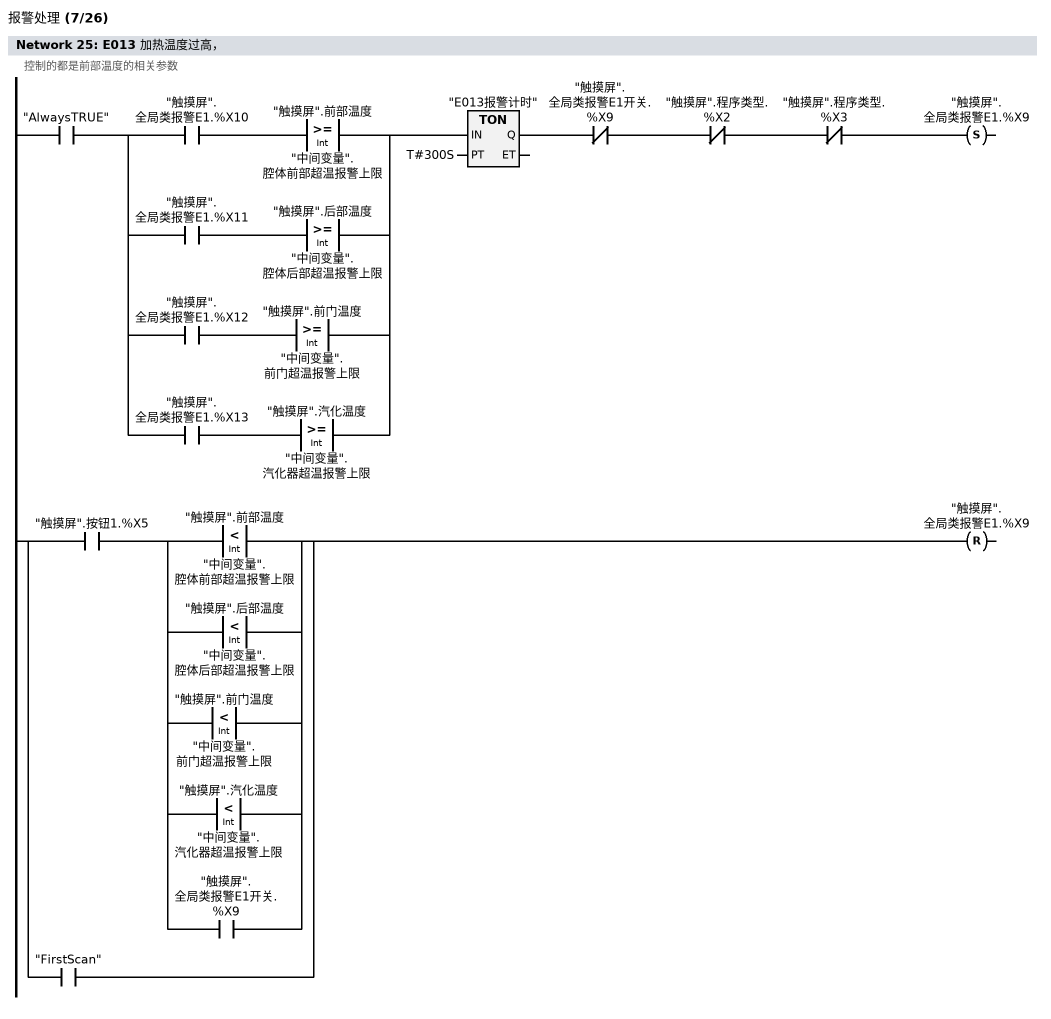
   "E013报警计时".TON(IN := "AlwaysTRUE" AND (("触摸屏".全局类报警E1.%X10 AND ("触摸屏".前部温度 >= "中间变量".腔体前部超温报警上限)) OR ("触摸屏".全局类报警E1.%X11 AND ("触摸屏".后部温度 >= "中间变量".腔体后部超温报警上限)) OR ("触摸屏".全局类报警E1.%X12 AND ("触摸屏".前门温度 >= "中间变量".前门超温报警上限)) OR ("触摸屏".全局类报警E1.%X13 AND ("触摸屏".汽化温度 >= "中间变量".汽化器超温报警上限))),
                  PT := T#300S);
   IF "E013报警计时".Q AND NOT "触摸屏".全局类报警E1开关.%X9 AND NOT "触摸屏".程序类型.%X2 AND NOT "触摸屏".程序类型.%X3 THEN
       "触摸屏".全局类报警E1.%X9 := TRUE;
   END_IF;
   IF ("触摸屏".按钮1.%X5 AND (("触摸屏".前部温度 < "中间变量".腔体前部超温报警上限) OR ("触摸屏".后部温度 < "中间变量".腔体后部超温报警上限) OR ("触摸屏".前门温度 < "中间变量".前门超温报警上限) OR ("触摸屏".汽化温度 < "中间变量".汽化器超温报警上限) OR "触摸屏".全局类报警E1开关.%X9)) OR "FirstScan" THEN
       "触摸屏".全局类报警E1.%X9 := FALSE;
   END_IF;
END_REGION

REGION Network 26: E014 加热系统异常，加热系统断电-脱扣器
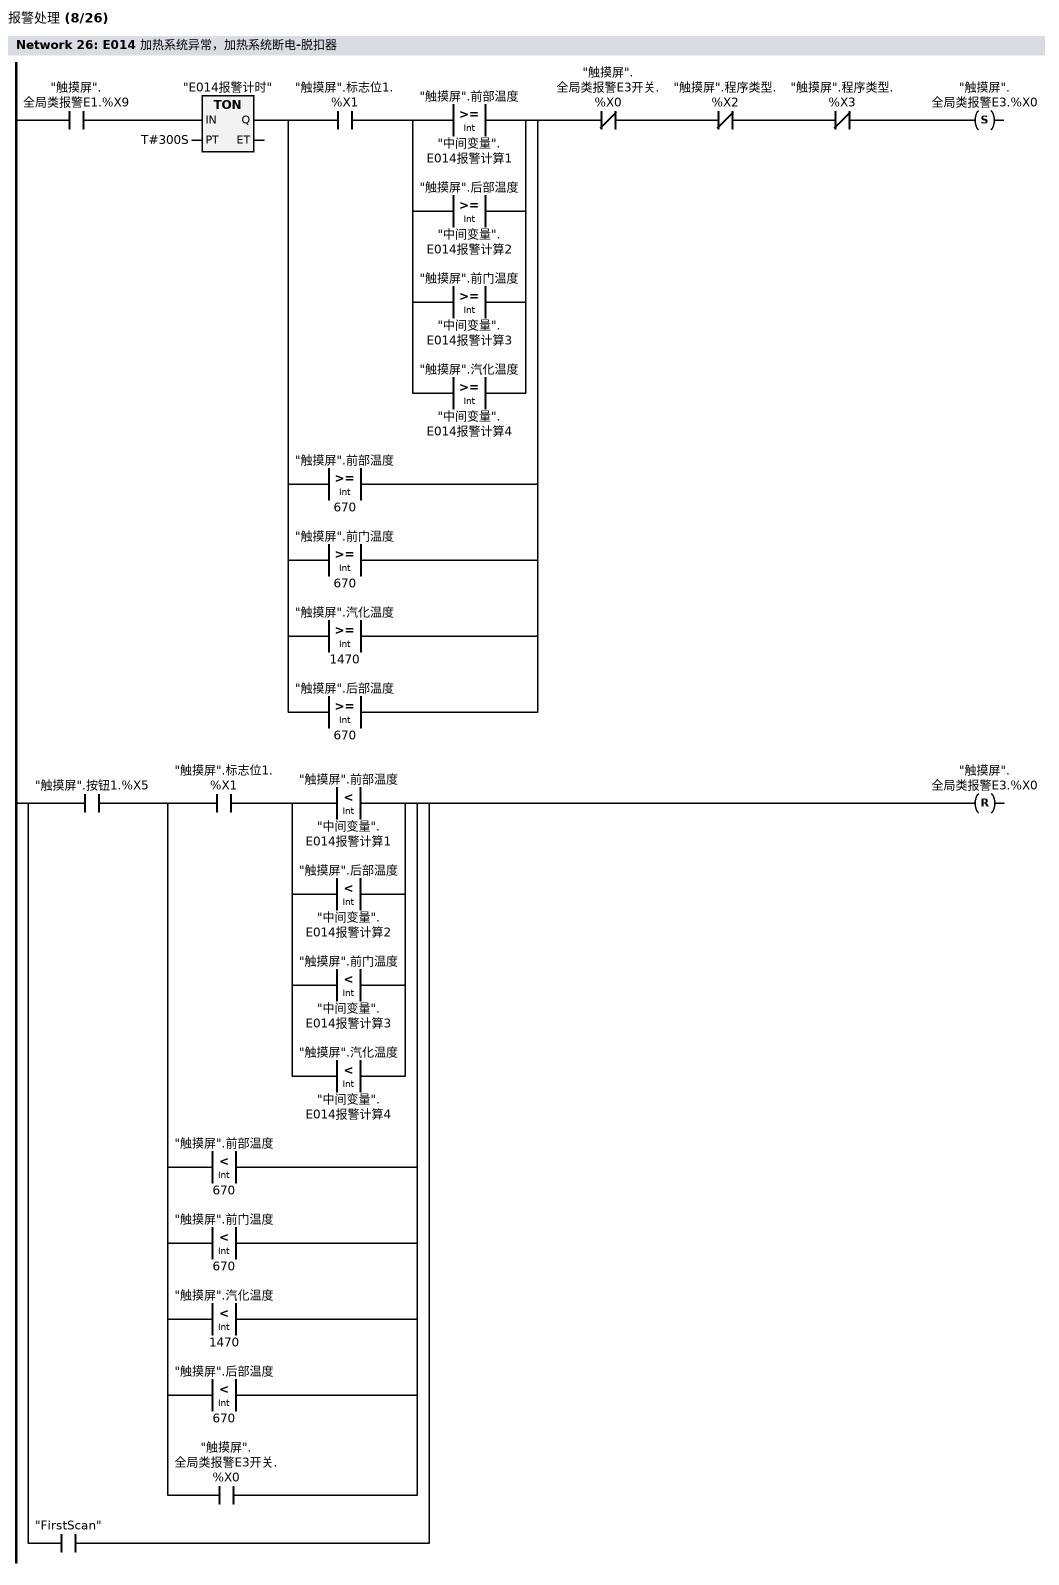
   "E014报警计时".TON(IN := "触摸屏".全局类报警E1.%X9, PT := T#300S);
   IF "E014报警计时".Q AND (("触摸屏".标志位1.%X1 AND (("触摸屏".前部温度 >= "中间变量".E014报警计算1) OR ("触摸屏".后部温度 >= "中间变量".E014报警计算2) OR ("触摸屏".前门温度 >= "中间变量".E014报警计算3) OR ("触摸屏".汽化温度 >= "中间变量".E014报警计算4))) OR ("触摸屏".前部温度 >= 670) OR ("触摸屏".前门温度 >= 670) OR ("触摸屏".汽化温度 >= 1470) OR ("触摸屏".后部温度 >= 670)) AND NOT "触摸屏".全局类报警E3开关.%X0 AND NOT "触摸屏".程序类型.%X2 AND NOT "触摸屏".程序类型.%X3 THEN
       "触摸屏".全局类报警E3.%X0 := TRUE;
   END_IF;
   IF ("触摸屏".按钮1.%X5 AND (("触摸屏".标志位1.%X1 AND (("触摸屏".前部温度 < "中间变量".E014报警计算1) OR ("触摸屏".后部温度 < "中间变量".E014报警计算2) OR ("触摸屏".前门温度 < "中间变量".E014报警计算3) OR ("触摸屏".汽化温度 < "中间变量".E014报警计算4))) OR ("触摸屏".前部温度 < 670) OR ("触摸屏".前门温度 < 670) OR ("触摸屏".汽化温度 < 1470) OR ("触摸屏".后部温度 < 670) OR "触摸屏".全局类报警E3开关.%X0)) OR "FirstScan" THEN
       "触摸屏".全局类报警E3.%X0 := FALSE;
   END_IF;
END_REGION

REGION Network 27: E015 腔体前部超温
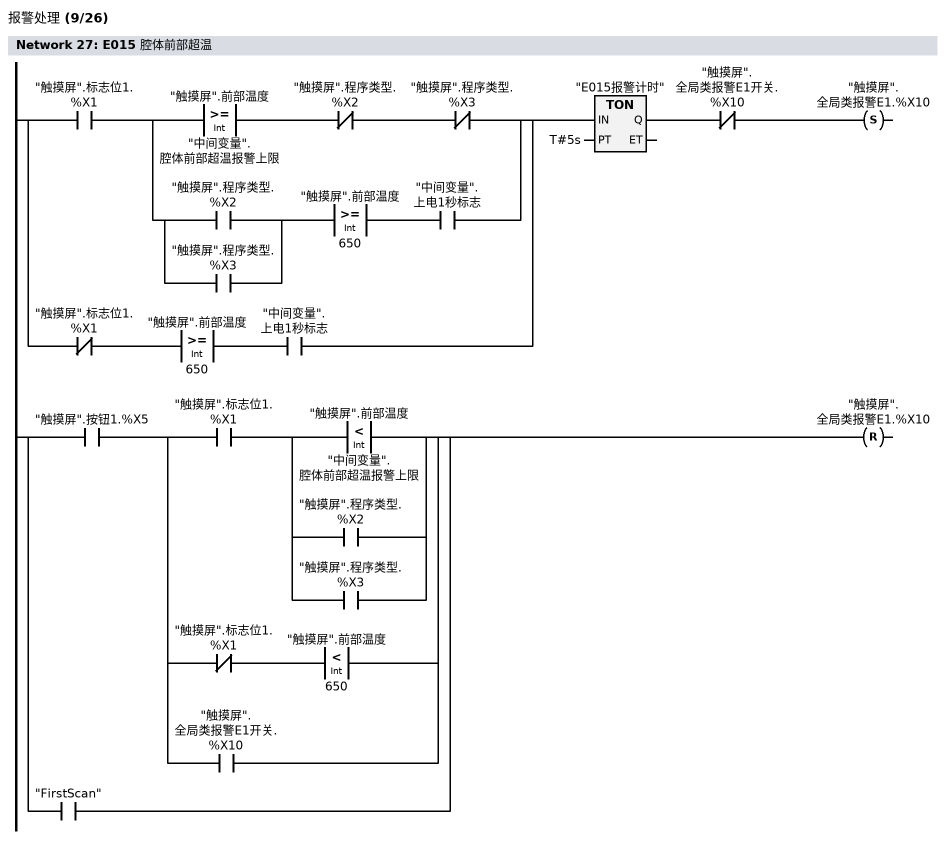
   "E015报警计时".TON(IN := ("触摸屏".标志位1.%X1 AND ((("触摸屏".前部温度 >= "中间变量".腔体前部超温报警上限) AND NOT "触摸屏".程序类型.%X2 AND NOT "触摸屏".程序类型.%X3) OR (("触摸屏".程序类型.%X2 OR "触摸屏".程序类型.%X3) AND ("触摸屏".前部温度 >= 650) AND "中间变量".上电1秒标志))) OR (NOT "触摸屏".标志位1.%X1 AND ("触摸屏".前部温度 >= 650) AND "中间变量".上电1秒标志),
                  PT := T#5s);
   IF "E015报警计时".Q AND NOT "触摸屏".全局类报警E1开关.%X10 THEN "触摸屏".全局类报警E1.%X10 := TRUE; END_IF;
   IF ("触摸屏".按钮1.%X5 AND (("触摸屏".标志位1.%X1 AND (("触摸屏".前部温度 < "中间变量".腔体前部超温报警上限) OR "触摸屏".程序类型.%X2 OR "触摸屏".程序类型.%X3)) OR (NOT "触摸屏".标志位1.%X1 AND ("触摸屏".前部温度 < 650)) OR "触摸屏".全局类报警E1开关.%X10)) OR "FirstScan" THEN
       "触摸屏".全局类报警E1.%X10 := FALSE;
   END_IF;
END_REGION

REGION Network 28: E016 腔体后部超温
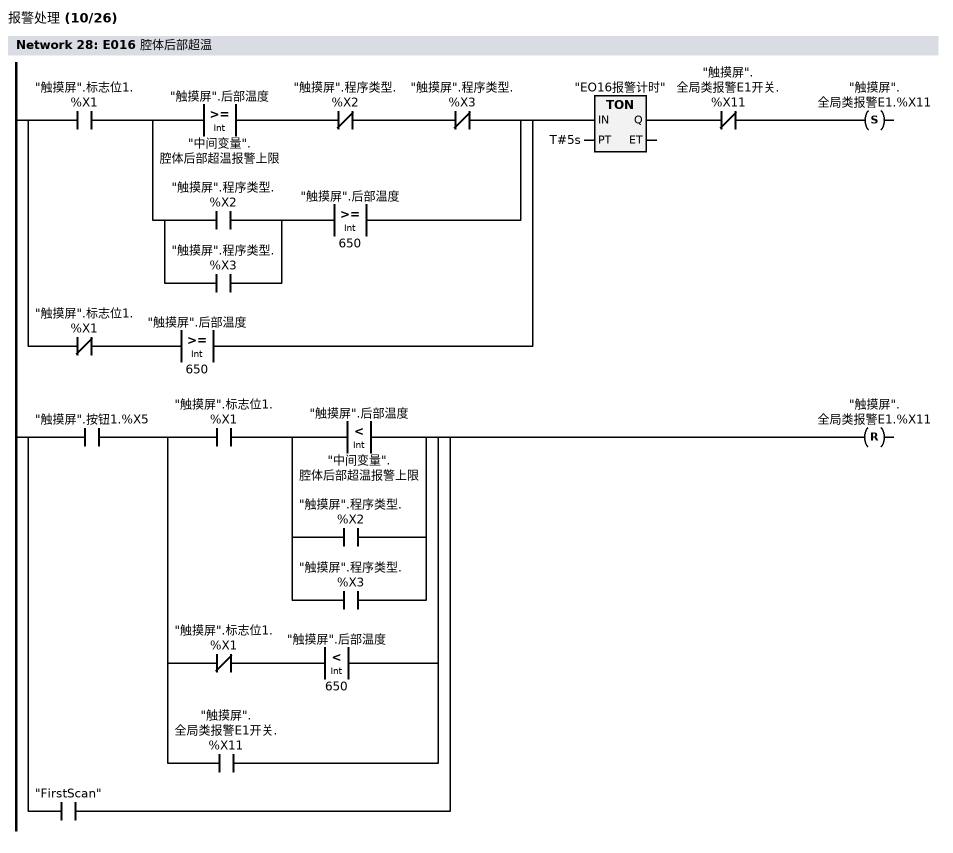
   "EO16报警计时".TON(IN := ("触摸屏".标志位1.%X1 AND ((("触摸屏".后部温度 >= "中间变量".腔体后部超温报警上限) AND NOT "触摸屏".程序类型.%X2 AND NOT "触摸屏".程序类型.%X3) OR (("触摸屏".程序类型.%X2 OR "触摸屏".程序类型.%X3) AND ("触摸屏".后部温度 >= 650)))) OR (NOT "触摸屏".标志位1.%X1 AND ("触摸屏".后部温度 >= 650)),
                  PT := T#5s);
   IF "EO16报警计时".Q AND NOT "触摸屏".全局类报警E1开关.%X11 THEN "触摸屏".全局类报警E1.%X11 := TRUE; END_IF;
   IF ("触摸屏".按钮1.%X5 AND (("触摸屏".标志位1.%X1 AND (("触摸屏".后部温度 < "中间变量".腔体后部超温报警上限) OR "触摸屏".程序类型.%X2 OR "触摸屏".程序类型.%X3)) OR (NOT "触摸屏".标志位1.%X1 AND ("触摸屏".后部温度 < 650)) OR "触摸屏".全局类报警E1开关.%X11)) OR "FirstScan" THEN
       "触摸屏".全局类报警E1.%X11 := FALSE;
   END_IF;
END_REGION

REGION Network 29: E017 门超温
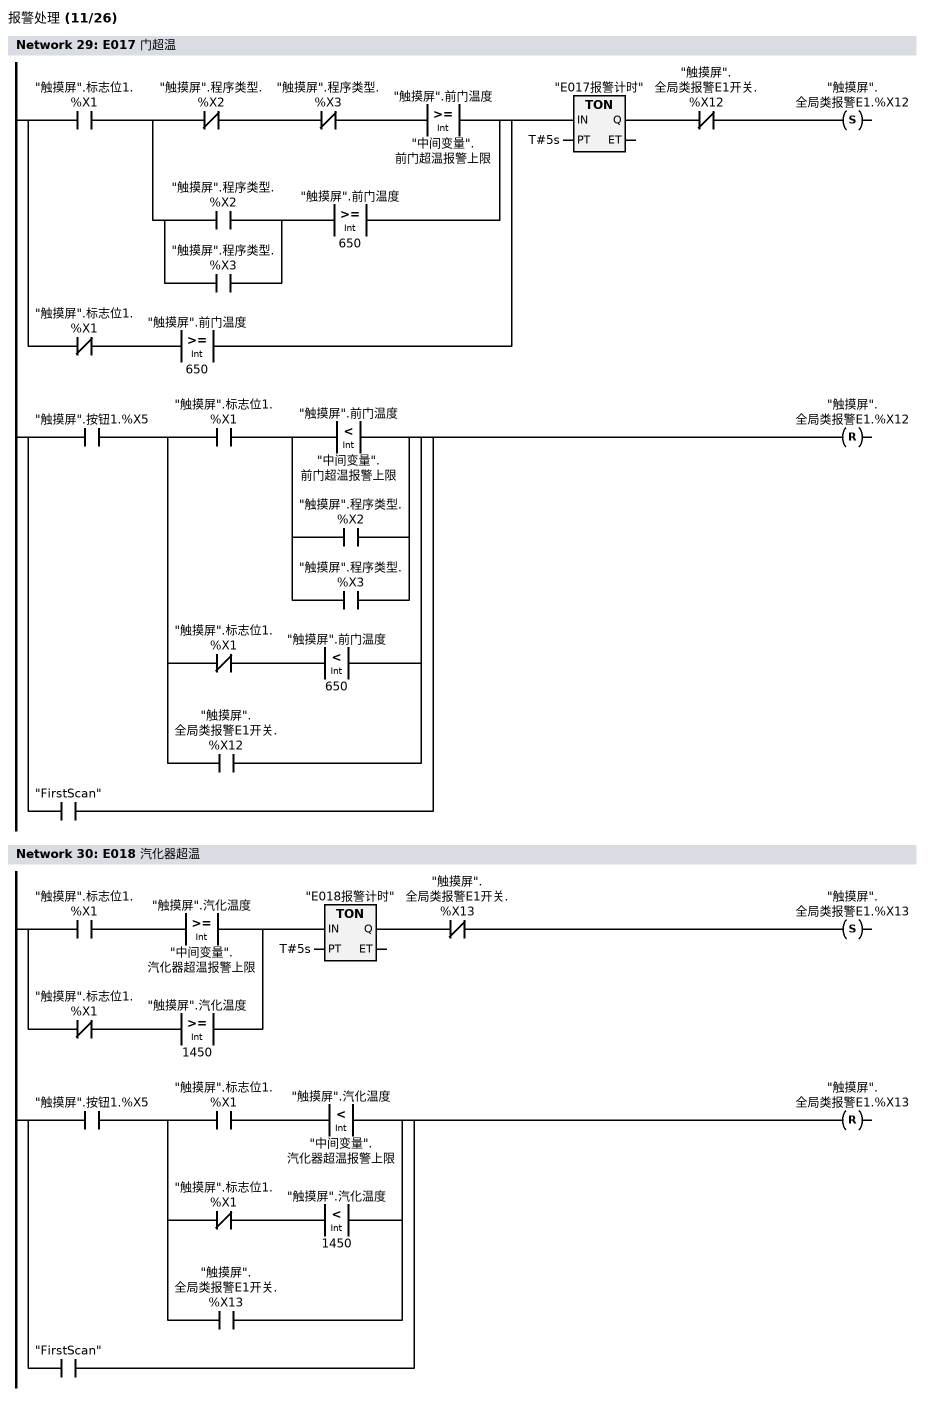
   "E017报警计时".TON(IN := ("触摸屏".标志位1.%X1 AND ((NOT "触摸屏".程序类型.%X2 AND NOT "触摸屏".程序类型.%X3 AND ("触摸屏".前门温度 >= "中间变量".前门超温报警上限)) OR (("触摸屏".程序类型.%X2 OR "触摸屏".程序类型.%X3) AND ("触摸屏".前门温度 >= 650)))) OR (NOT "触摸屏".标志位1.%X1 AND ("触摸屏".前门温度 >= 650)),
                  PT := T#5s);
   IF "E017报警计时".Q AND NOT "触摸屏".全局类报警E1开关.%X12 THEN "触摸屏".全局类报警E1.%X12 := TRUE; END_IF;
   IF ("触摸屏".按钮1.%X5 AND (("触摸屏".标志位1.%X1 AND (("触摸屏".前门温度 < "中间变量".前门超温报警上限) OR "触摸屏".程序类型.%X2 OR "触摸屏".程序类型.%X3)) OR (NOT "触摸屏".标志位1.%X1 AND ("触摸屏".前门温度 < 650)) OR "触摸屏".全局类报警E1开关.%X12)) OR "FirstScan" THEN
       "触摸屏".全局类报警E1.%X12 := FALSE;
   END_IF;
END_REGION

REGION Network 30: E018 汽化器超温
   "E018报警计时".TON(IN := ("触摸屏".标志位1.%X1 AND ("触摸屏".汽化温度 >= "中间变量".汽化器超温报警上限)) OR (NOT "触摸屏".标志位1.%X1 AND ("触摸屏".汽化温度 >= 1450)),
                  PT := T#5s);
   IF "E018报警计时".Q AND NOT "触摸屏".全局类报警E1开关.%X13 THEN "触摸屏".全局类报警E1.%X13 := TRUE; END_IF;
   IF ("触摸屏".按钮1.%X5 AND (("触摸屏".标志位1.%X1 AND ("触摸屏".汽化温度 < "中间变量".汽化器超温报警上限)) OR (NOT "触摸屏".标志位1.%X1 AND ("触摸屏".汽化温度 < 1450)) OR "触摸屏".全局类报警E1开关.%X13)) OR "FirstScan" THEN
       "触摸屏".全局类报警E1.%X13 := FALSE;
   END_IF;
END_REGION

REGION Network 31: E019 内室温度过高
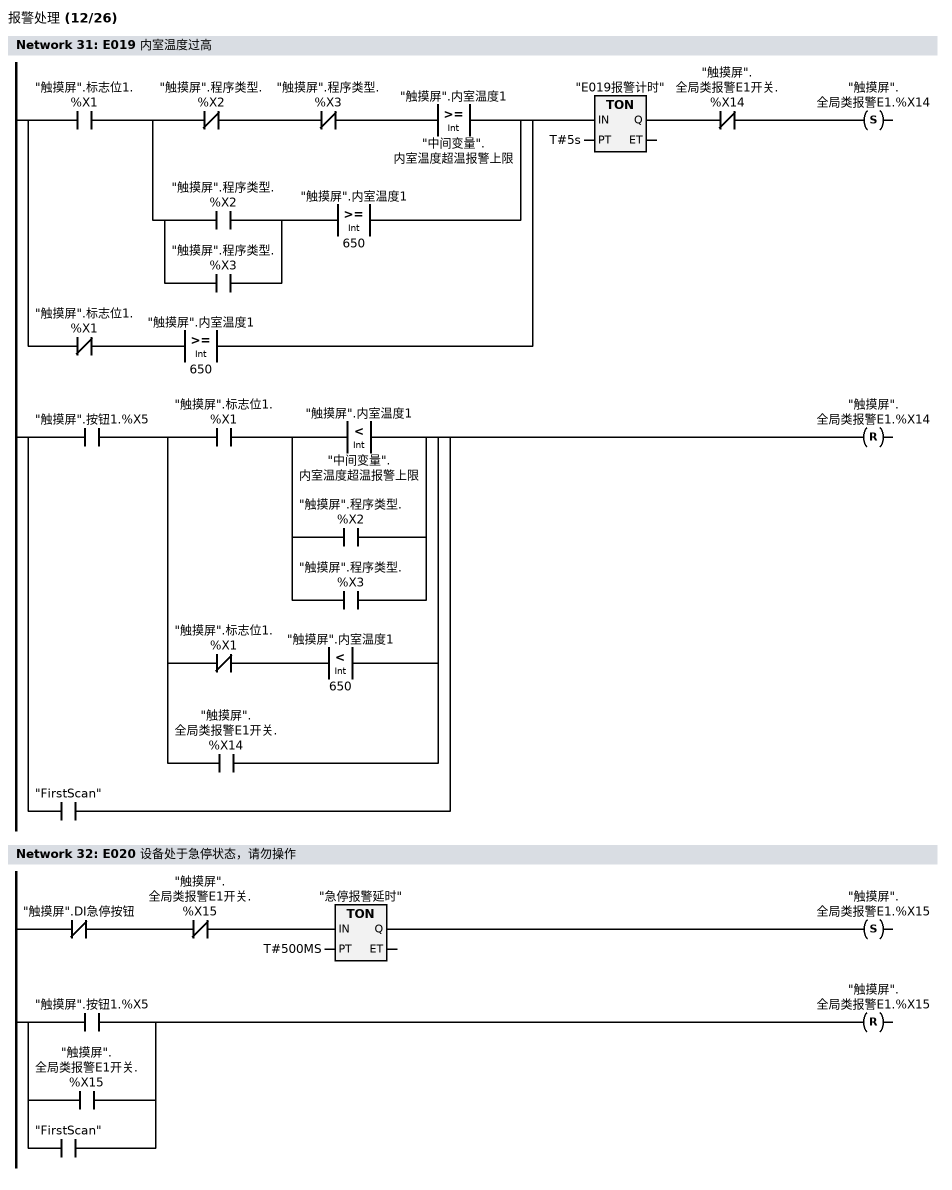
   "E019报警计时".TON(IN := ("触摸屏".标志位1.%X1 AND ((NOT "触摸屏".程序类型.%X2 AND NOT "触摸屏".程序类型.%X3 AND ("触摸屏".内室温度1 >= "中间变量".内室温度超温报警上限)) OR (("触摸屏".程序类型.%X2 OR "触摸屏".程序类型.%X3) AND ("触摸屏".内室温度1 >= 650)))) OR (NOT "触摸屏".标志位1.%X1 AND ("触摸屏".内室温度1 >= 650)),
                  PT := T#5s);
   IF "E019报警计时".Q AND NOT "触摸屏".全局类报警E1开关.%X14 THEN "触摸屏".全局类报警E1.%X14 := TRUE; END_IF;
   IF ("触摸屏".按钮1.%X5 AND (("触摸屏".标志位1.%X1 AND (("触摸屏".内室温度1 < "中间变量".内室温度超温报警上限) OR "触摸屏".程序类型.%X2 OR "触摸屏".程序类型.%X3)) OR (NOT "触摸屏".标志位1.%X1 AND ("触摸屏".内室温度1 < 650)) OR "触摸屏".全局类报警E1开关.%X14)) OR "FirstScan" THEN
       "触摸屏".全局类报警E1.%X14 := FALSE;
   END_IF;
END_REGION

REGION Network 32: E020 设备处于急停状态，请勿操作
   "急停报警延时".TON(IN := NOT "触摸屏".DI急停按钮 AND NOT "触摸屏".全局类报警E1开关.%X15, PT := T#500MS);
   IF "急停报警延时".Q THEN "触摸屏".全局类报警E1.%X15 := TRUE; END_IF;
   IF "触摸屏".按钮1.%X5 OR "触摸屏".全局类报警E1开关.%X15 OR "FirstScan" THEN "触摸屏".全局类报警E1.%X15 := FALSE; END_IF;
END_REGION

REGION Network 33: E021灭菌器与尾气处理器通讯故障
   // 带尾气处理器的设备   通讯超时60秒 我们认为通讯故障
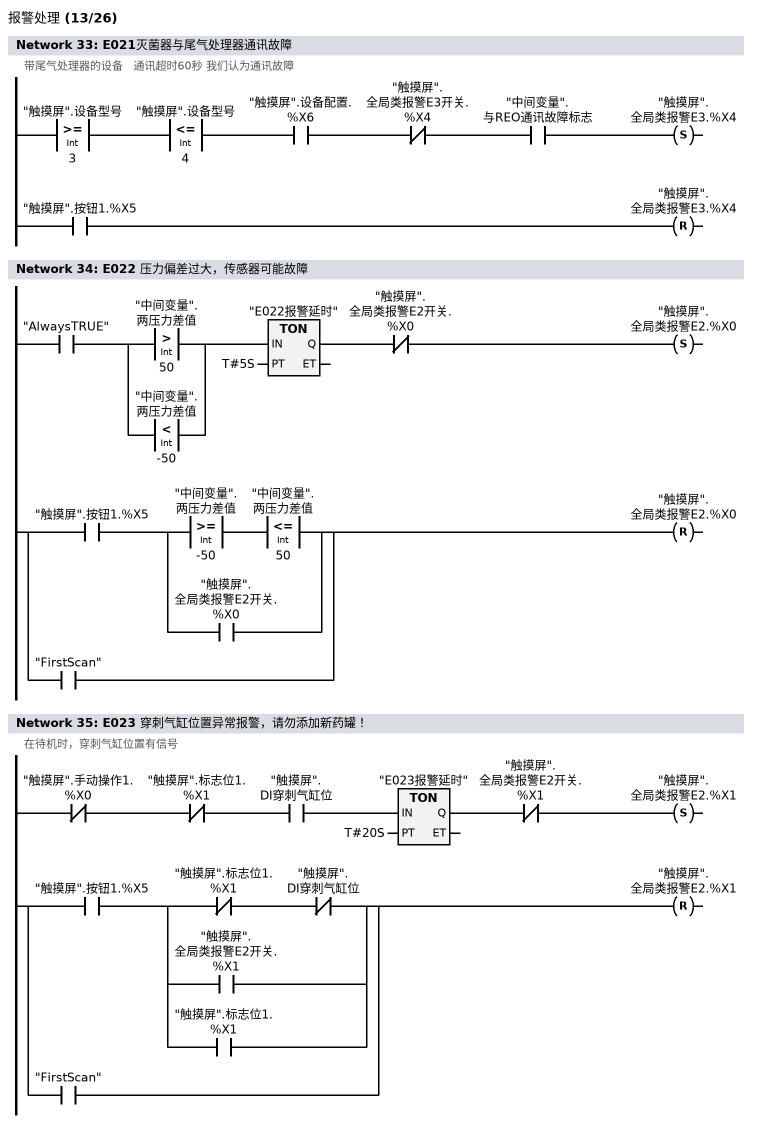
   RUNG wire#powerrail
      { S7_Templates := "SrcType := Int" } GE_Contact(in1 := "触摸屏".设备型号, in2 := 3)
      { S7_Templates := "SrcType := Int" } LE_Contact(in1 := "触摸屏".设备型号, in2 := 4)
      Contact( "触摸屏".设备配置.%X6 )
      I_Contact( "触摸屏".全局类报警E3开关.%X4 )
      Contact( "中间变量".与REO通讯故障标志 )
      S_Coil( "触摸屏".全局类报警E3.%X4 )
   END_RUNG
   RUNG wire#powerrail
      Contact( "触摸屏".按钮1.%X5 )
      R_Coil( "触摸屏".全局类报警E3.%X4 )
   END_RUNG
   // the same network as SCL:
   IF ("触摸屏".设备型号 >= 3) AND ("触摸屏".设备型号 <= 4) AND "触摸屏".设备配置.%X6 AND NOT "触摸屏".全局类报警E3开关.%X4 AND "中间变量".与REO通讯故障标志 THEN
       "触摸屏".全局类报警E3.%X4 := TRUE;
   END_IF;
   IF "触摸屏".按钮1.%X5 THEN "触摸屏".全局类报警E3.%X4 := FALSE; END_IF;
END_REGION

REGION Network 34: E022 压力偏差过大，传感器可能故障
   "E022报警延时".TON(IN := "AlwaysTRUE" AND (("中间变量".两压力差值 > 50) OR ("中间变量".两压力差值 < (-50))), PT := T#5S);
   IF "E022报警延时".Q AND NOT "触摸屏".全局类报警E2开关.%X0 THEN "触摸屏".全局类报警E2.%X0 := TRUE; END_IF;
   IF ("触摸屏".按钮1.%X5 AND ((("中间变量".两压力差值 >= (-50)) AND ("中间变量".两压力差值 <= 50)) OR "触摸屏".全局类报警E2开关.%X0)) OR "FirstScan" THEN
       "触摸屏".全局类报警E2.%X0 := FALSE;
   END_IF;
END_REGION

REGION Network 35: E023 穿刺气缸位置异常报警，请勿添加新药罐！
   // 在待机时，穿刺气缸位置有信号
   "E023报警延时".TON(IN := NOT "触摸屏".手动操作1.%X0 AND NOT "触摸屏".标志位1.%X1 AND "触摸屏".DI穿刺气缸位, PT := T#20S);
   IF "E023报警延时".Q AND NOT "触摸屏".全局类报警E2开关.%X1 THEN "触摸屏".全局类报警E2.%X1 := TRUE; END_IF;
   IF ("触摸屏".按钮1.%X5 AND ((NOT "触摸屏".标志位1.%X1 AND NOT "触摸屏".DI穿刺气缸位) OR "触摸屏".全局类报警E2开关.%X1 OR "触摸屏".标志位1.%X1)) OR "FirstScan" THEN
       "触摸屏".全局类报警E2.%X1 := FALSE;
   END_IF;
END_REGION

REGION Network 36: E024舱体前部温度升温超时
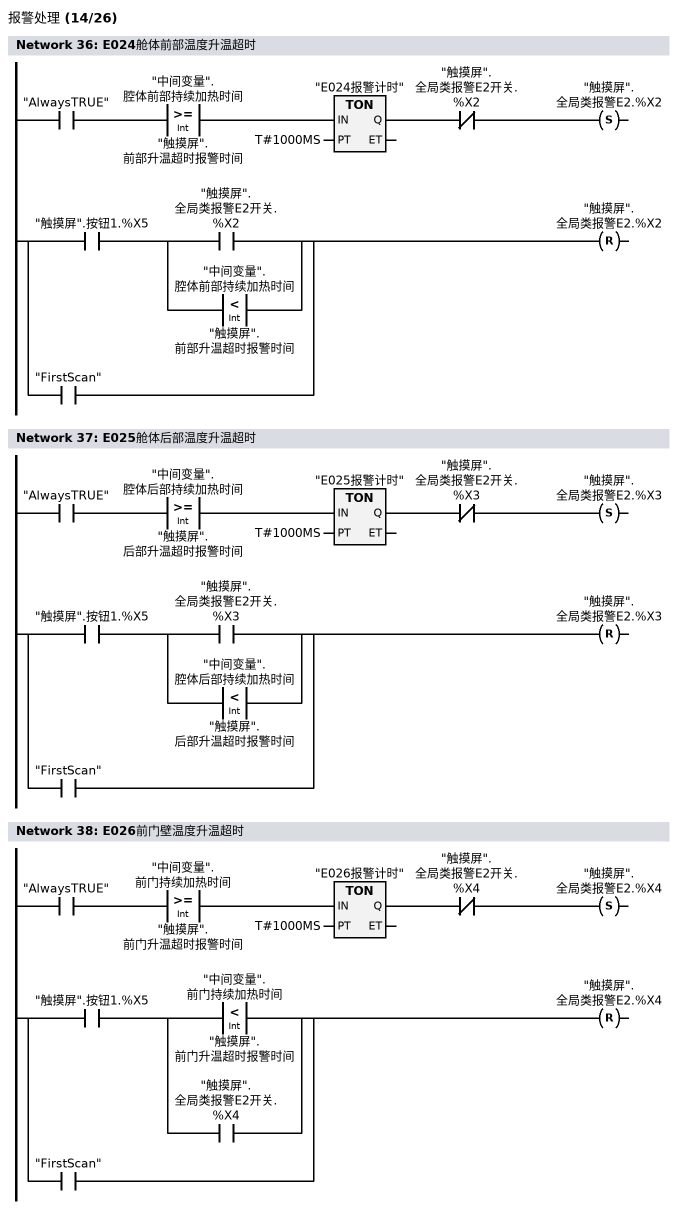
   "E024报警计时".TON(IN := "AlwaysTRUE" AND ("中间变量".腔体前部持续加热时间 >= "触摸屏".前部升温超时报警时间), PT := T#1000MS);
   IF "E024报警计时".Q AND NOT "触摸屏".全局类报警E2开关.%X2 THEN "触摸屏".全局类报警E2.%X2 := TRUE; END_IF;
   IF ("触摸屏".按钮1.%X5 AND ("触摸屏".全局类报警E2开关.%X2 OR ("中间变量".腔体前部持续加热时间 < "触摸屏".前部升温超时报警时间))) OR "FirstScan" THEN
       "触摸屏".全局类报警E2.%X2 := FALSE;
   END_IF;
END_REGION

REGION Network 37: E025舱体后部温度升温超时
   "E025报警计时".TON(IN := "AlwaysTRUE" AND ("中间变量".腔体后部持续加热时间 >= "触摸屏".后部升温超时报警时间), PT := T#1000MS);
   IF "E025报警计时".Q AND NOT "触摸屏".全局类报警E2开关.%X3 THEN "触摸屏".全局类报警E2.%X3 := TRUE; END_IF;
   IF ("触摸屏".按钮1.%X5 AND ("触摸屏".全局类报警E2开关.%X3 OR ("中间变量".腔体后部持续加热时间 < "触摸屏".后部升温超时报警时间))) OR "FirstScan" THEN
       "触摸屏".全局类报警E2.%X3 := FALSE;
   END_IF;
END_REGION

REGION Network 38: E026前门壁温度升温超时
   "E026报警计时".TON(IN := "AlwaysTRUE" AND ("中间变量".前门持续加热时间 >= "触摸屏".前门升温超时报警时间), PT := T#1000MS);
   IF "E026报警计时".Q AND NOT "触摸屏".全局类报警E2开关.%X4 THEN "触摸屏".全局类报警E2.%X4 := TRUE; END_IF;
   IF ("触摸屏".按钮1.%X5 AND (("中间变量".前门持续加热时间 < "触摸屏".前门升温超时报警时间) OR "触摸屏".全局类报警E2开关.%X4)) OR "FirstScan" THEN
       "触摸屏".全局类报警E2.%X4 := FALSE;
   END_IF;
END_REGION

REGION Network 39: E027汽化器温度升温超时
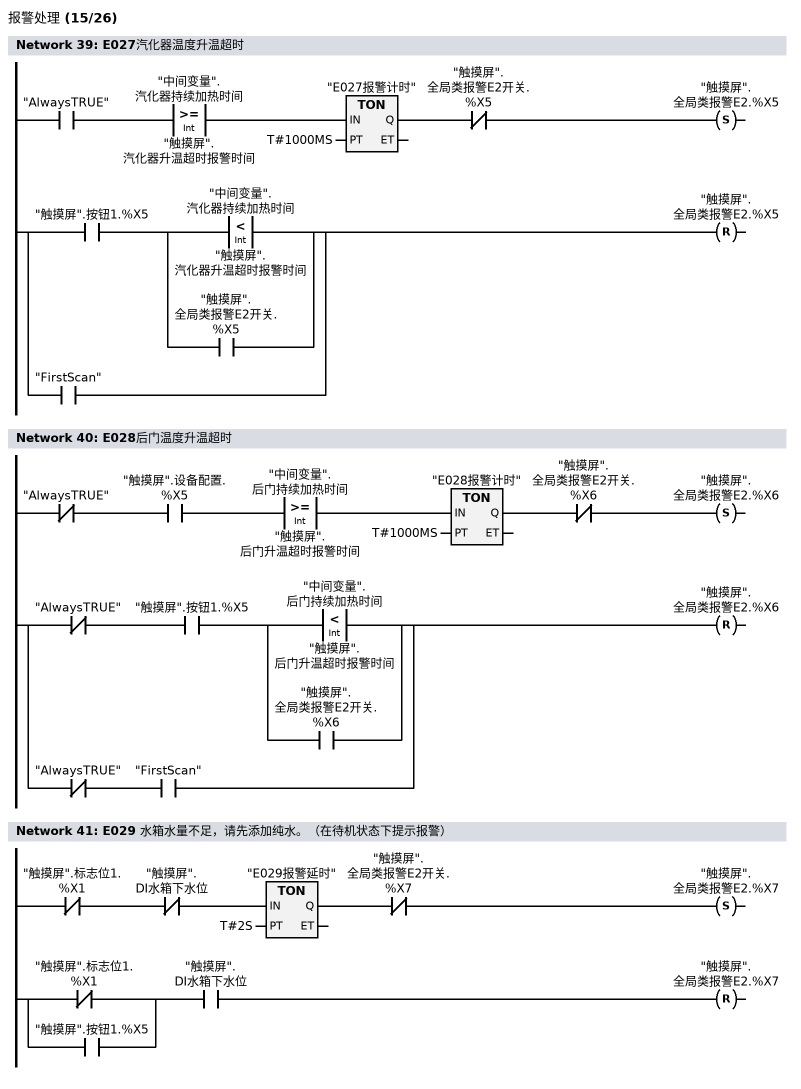
   "E027报警计时".TON(IN := "AlwaysTRUE" AND ("中间变量".汽化器持续加热时间 >= "触摸屏".汽化器升温超时报警时间), PT := T#1000MS);
   IF "E027报警计时".Q AND NOT "触摸屏".全局类报警E2开关.%X5 THEN "触摸屏".全局类报警E2.%X5 := TRUE; END_IF;
   IF ("触摸屏".按钮1.%X5 AND (("中间变量".汽化器持续加热时间 < "触摸屏".汽化器升温超时报警时间) OR "触摸屏".全局类报警E2开关.%X5)) OR "FirstScan" THEN
       "触摸屏".全局类报警E2.%X5 := FALSE;
   END_IF;
END_REGION

REGION Network 40: E028后门温度升温超时
   "E028报警计时".TON(IN := NOT "AlwaysTRUE" AND "触摸屏".设备配置.%X5 AND ("中间变量".后门持续加热时间 >= "触摸屏".后门升温超时报警时间),
                  PT := T#1000MS);
   IF "E028报警计时".Q AND NOT "触摸屏".全局类报警E2开关.%X6 THEN "触摸屏".全局类报警E2.%X6 := TRUE; END_IF;
   IF (NOT "AlwaysTRUE" AND "触摸屏".按钮1.%X5 AND (("中间变量".后门持续加热时间 < "触摸屏".后门升温超时报警时间) OR "触摸屏".全局类报警E2开关.%X6)) OR (NOT "AlwaysTRUE" AND "FirstScan") THEN
       "触摸屏".全局类报警E2.%X6 := FALSE;
   END_IF;
END_REGION

REGION Network 41: E029 水箱水量不足，请先添加纯水。（在待机状态下提示报警）
   "E029报警延时".TON(IN := NOT "触摸屏".标志位1.%X1 AND NOT "触摸屏".DI水箱下水位, PT := T#2S);
   IF "E029报警延时".Q AND NOT "触摸屏".全局类报警E2开关.%X7 THEN "触摸屏".全局类报警E2.%X7 := TRUE; END_IF;
   IF (NOT "触摸屏".标志位1.%X1 OR "触摸屏".按钮1.%X5) AND "触摸屏".DI水箱下水位 THEN "触摸屏".全局类报警E2.%X7 := FALSE; END_IF;
END_REGION

REGION Network 42: E030催化前温度传感器故障！
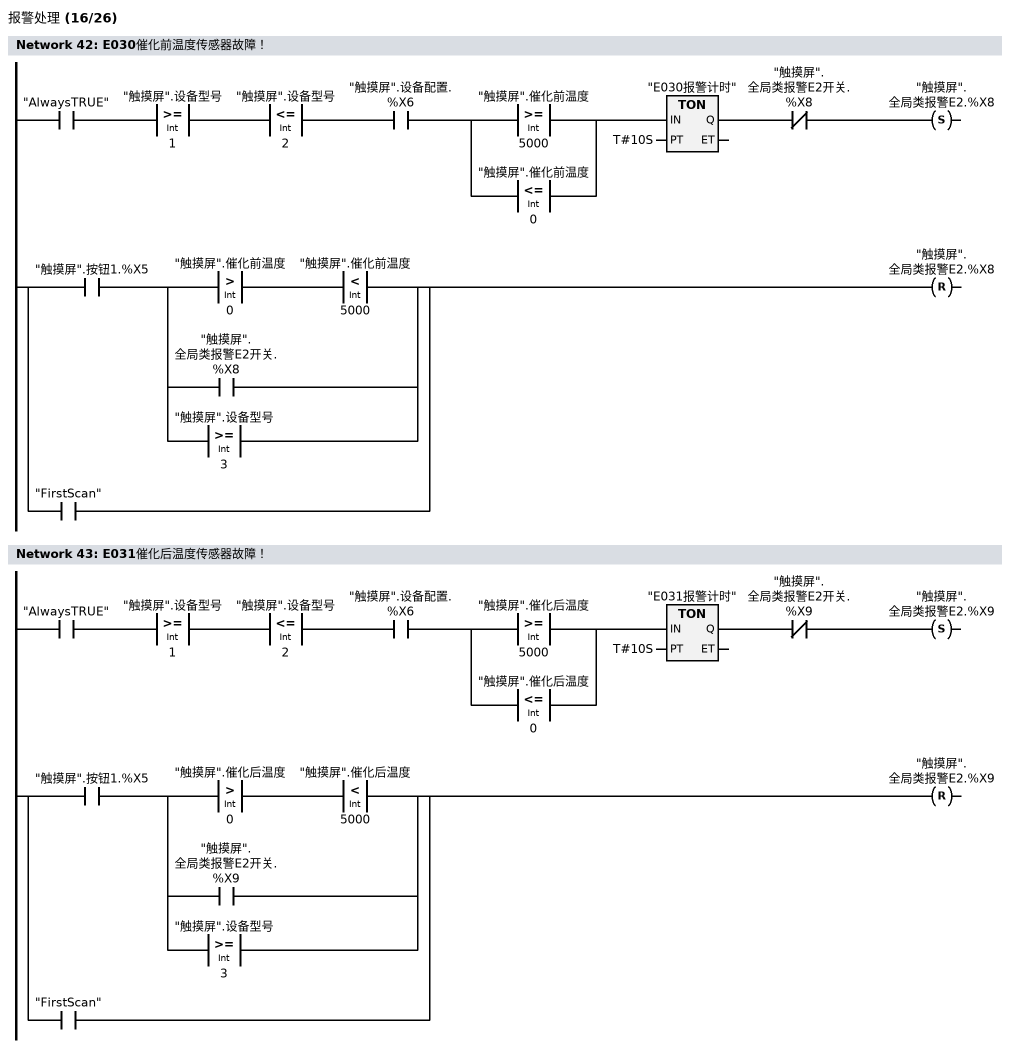
   "E030报警计时".TON(IN := "AlwaysTRUE" AND ("触摸屏".设备型号 >= 1) AND ("触摸屏".设备型号 <= 2) AND "触摸屏".设备配置.%X6 AND (("触摸屏".催化前温度 >= 5000) OR ("触摸屏".催化前温度 <= 0)),
                  PT := T#10S);
   IF "E030报警计时".Q AND NOT "触摸屏".全局类报警E2开关.%X8 THEN "触摸屏".全局类报警E2.%X8 := TRUE; END_IF;
   IF ("触摸屏".按钮1.%X5 AND ((("触摸屏".催化前温度 > 0) AND ("触摸屏".催化前温度 < 5000)) OR "触摸屏".全局类报警E2开关.%X8 OR ("触摸屏".设备型号 >= 3))) OR "FirstScan" THEN
       "触摸屏".全局类报警E2.%X8 := FALSE;
   END_IF;
END_REGION

REGION Network 43: E031催化后温度传感器故障！
   "E031报警计时".TON(IN := "AlwaysTRUE" AND ("触摸屏".设备型号 >= 1) AND ("触摸屏".设备型号 <= 2) AND "触摸屏".设备配置.%X6 AND (("触摸屏".催化后温度 >= 5000) OR ("触摸屏".催化后温度 <= 0)),
                  PT := T#10S);
   IF "E031报警计时".Q AND NOT "触摸屏".全局类报警E2开关.%X9 THEN "触摸屏".全局类报警E2.%X9 := TRUE; END_IF;
   IF ("触摸屏".按钮1.%X5 AND ((("触摸屏".催化后温度 > 0) AND ("触摸屏".催化后温度 < 5000)) OR "触摸屏".全局类报警E2开关.%X9 OR ("触摸屏".设备型号 >= 3))) OR "FirstScan" THEN
       "触摸屏".全局类报警E2.%X9 := FALSE;
   END_IF;
END_REGION

REGION Network 44: E032后门温度传感器故障！
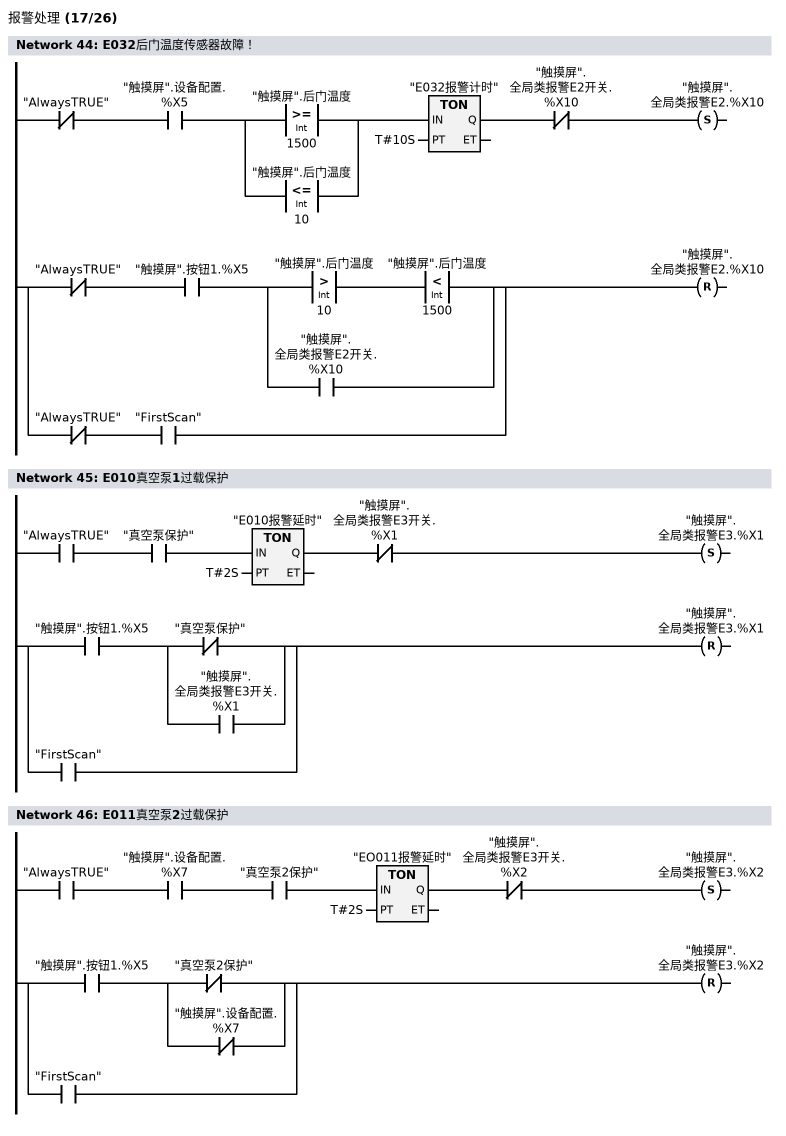
   "E032报警计时".TON(IN := NOT "AlwaysTRUE" AND "触摸屏".设备配置.%X5 AND (("触摸屏".后门温度 >= 1500) OR ("触摸屏".后门温度 <= 10)),
                  PT := T#10S);
   IF "E032报警计时".Q AND NOT "触摸屏".全局类报警E2开关.%X10 THEN "触摸屏".全局类报警E2.%X10 := TRUE; END_IF;
   IF (NOT "AlwaysTRUE" AND "触摸屏".按钮1.%X5 AND ((("触摸屏".后门温度 > 10) AND ("触摸屏".后门温度 < 1500)) OR "触摸屏".全局类报警E2开关.%X10)) OR (NOT "AlwaysTRUE" AND "FirstScan") THEN
       "触摸屏".全局类报警E2.%X10 := FALSE;
   END_IF;
END_REGION

REGION Network 45: E010真空泵1过载保护
   "E010报警延时".TON(IN := "AlwaysTRUE" AND "真空泵保护", PT := T#2S);
   IF "E010报警延时".Q AND NOT "触摸屏".全局类报警E3开关.%X1 THEN "触摸屏".全局类报警E3.%X1 := TRUE; END_IF;
   IF ("触摸屏".按钮1.%X5 AND (NOT "真空泵保护" OR "触摸屏".全局类报警E3开关.%X1)) OR "FirstScan" THEN
       "触摸屏".全局类报警E3.%X1 := FALSE;
   END_IF;
END_REGION

REGION Network 46: E011真空泵2过载保护
   "EO011报警延时".TON(IN := "AlwaysTRUE" AND "触摸屏".设备配置.%X7 AND "真空泵2保护", PT := T#2S);
   IF "EO011报警延时".Q AND NOT "触摸屏".全局类报警E3开关.%X2 THEN "触摸屏".全局类报警E3.%X2 := TRUE; END_IF;
   IF ("触摸屏".按钮1.%X5 AND (NOT "真空泵2保护" OR NOT "触摸屏".设备配置.%X7)) OR "FirstScan" THEN
       "触摸屏".全局类报警E3.%X2 := FALSE;
   END_IF;
END_REGION

REGION Network 47: E012空压机过载保护
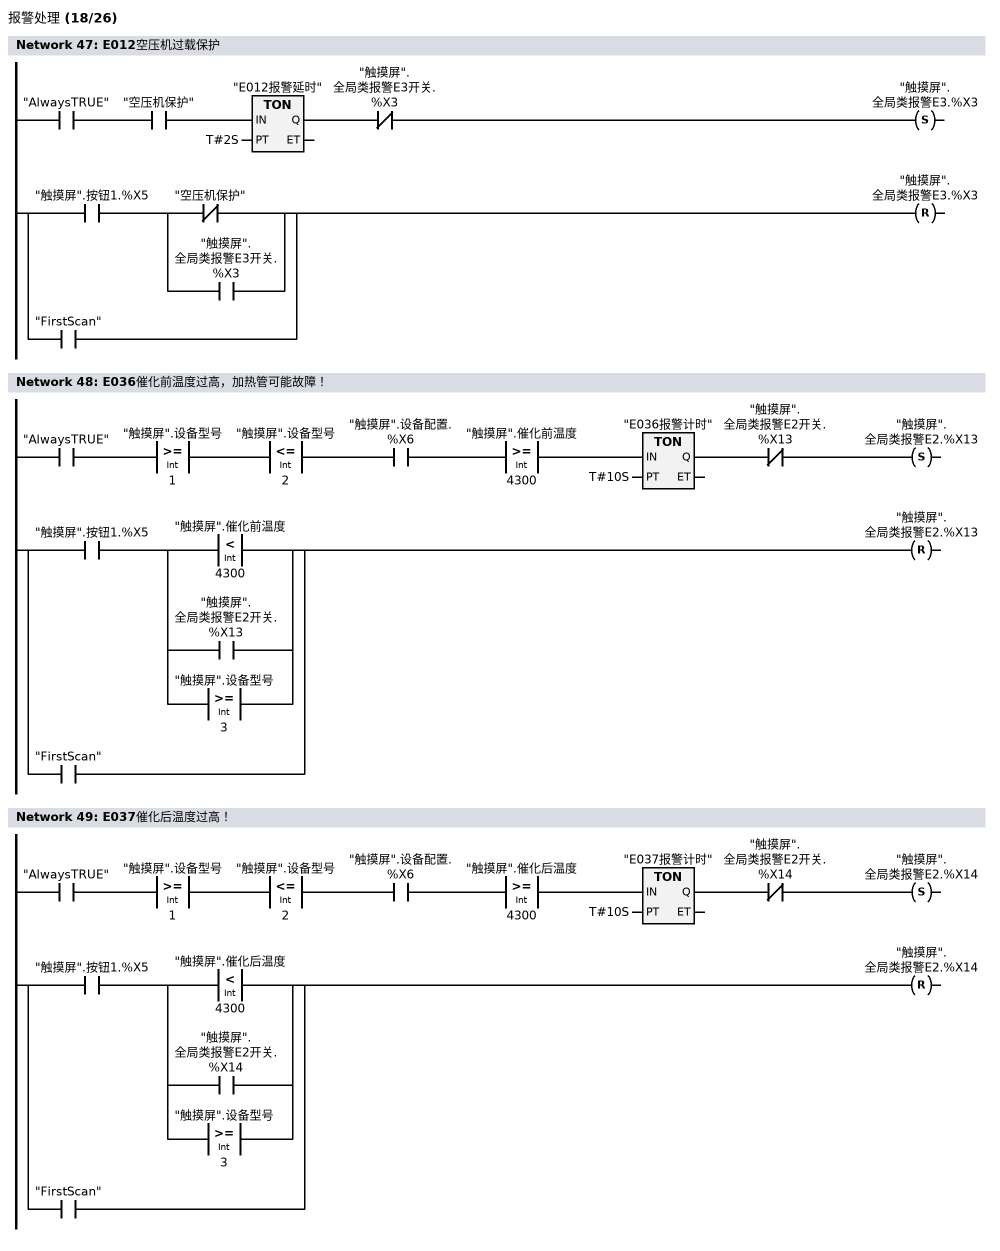
   "E012报警延时".TON(IN := "AlwaysTRUE" AND "空压机保护", PT := T#2S);
   IF "E012报警延时".Q AND NOT "触摸屏".全局类报警E3开关.%X3 THEN "触摸屏".全局类报警E3.%X3 := TRUE; END_IF;
   IF ("触摸屏".按钮1.%X5 AND (NOT "空压机保护" OR "触摸屏".全局类报警E3开关.%X3)) OR "FirstScan" THEN
       "触摸屏".全局类报警E3.%X3 := FALSE;
   END_IF;
END_REGION

REGION Network 48: E036催化前温度过高，加热管可能故障！
   "E036报警计时".TON(IN := "AlwaysTRUE" AND ("触摸屏".设备型号 >= 1) AND ("触摸屏".设备型号 <= 2) AND "触摸屏".设备配置.%X6 AND ("触摸屏".催化前温度 >= 4300),
                  PT := T#10S);
   IF "E036报警计时".Q AND NOT "触摸屏".全局类报警E2开关.%X13 THEN "触摸屏".全局类报警E2.%X13 := TRUE; END_IF;
   IF ("触摸屏".按钮1.%X5 AND (("触摸屏".催化前温度 < 4300) OR "触摸屏".全局类报警E2开关.%X13 OR ("触摸屏".设备型号 >= 3))) OR "FirstScan" THEN
       "触摸屏".全局类报警E2.%X13 := FALSE;
   END_IF;
END_REGION

REGION Network 49: E037催化后温度过高！
   "E037报警计时".TON(IN := "AlwaysTRUE" AND ("触摸屏".设备型号 >= 1) AND ("触摸屏".设备型号 <= 2) AND "触摸屏".设备配置.%X6 AND ("触摸屏".催化后温度 >= 4300),
                  PT := T#10S);
   IF "E037报警计时".Q AND NOT "触摸屏".全局类报警E2开关.%X14 THEN "触摸屏".全局类报警E2.%X14 := TRUE; END_IF;
   IF ("触摸屏".按钮1.%X5 AND (("触摸屏".催化后温度 < 4300) OR "触摸屏".全局类报警E2开关.%X14 OR ("触摸屏".设备型号 >= 3))) OR "FirstScan" THEN
       "触摸屏".全局类报警E2.%X14 := FALSE;
   END_IF;
END_REGION

REGION Network 50: E038催化加热升温超时！
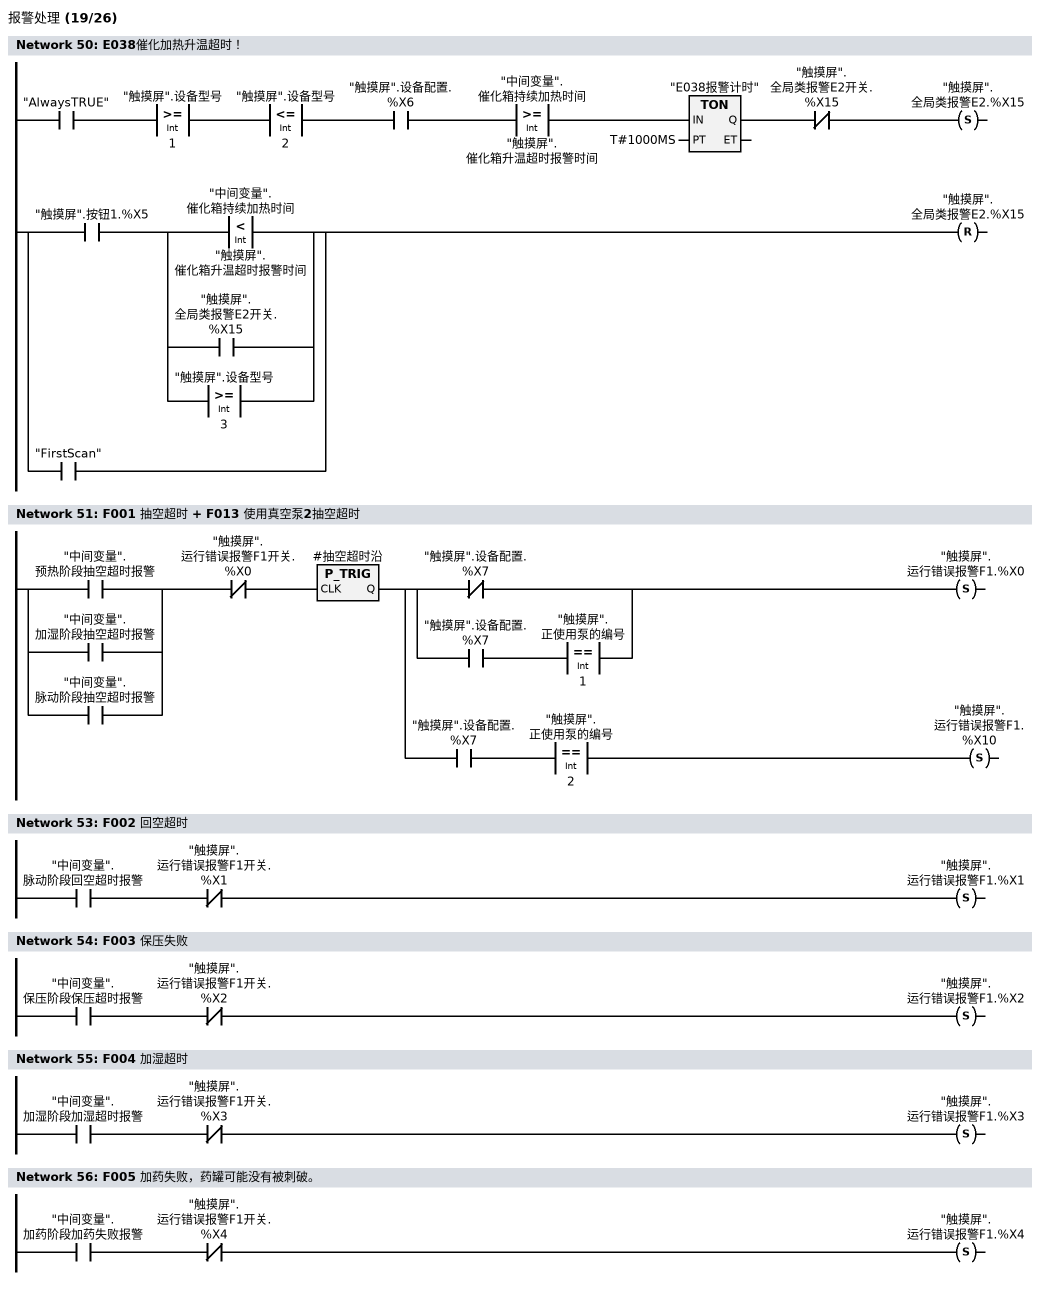
   "E038报警计时".TON(IN := "AlwaysTRUE" AND ("触摸屏".设备型号 >= 1) AND ("触摸屏".设备型号 <= 2) AND "触摸屏".设备配置.%X6 AND ("中间变量".催化箱持续加热时间 >= "触摸屏".催化箱升温超时报警时间),
                  PT := T#1000MS);
   IF "E038报警计时".Q AND NOT "触摸屏".全局类报警E2开关.%X15 THEN "触摸屏".全局类报警E2.%X15 := TRUE; END_IF;
   IF ("触摸屏".按钮1.%X5 AND (("中间变量".催化箱持续加热时间 < "触摸屏".催化箱升温超时报警时间) OR "触摸屏".全局类报警E2开关.%X15 OR ("触摸屏".设备型号 >= 3))) OR "FirstScan" THEN
       "触摸屏".全局类报警E2.%X15 := FALSE;
   END_IF;
END_REGION

REGION Network 51: F001 抽空超时 + F013 使用真空泵2抽空超时
   RUNG wire#powerrail
      Contact( "中间变量".预热阶段抽空超时报警 )
      wire#w1
      I_Contact( "触摸屏".运行错误报警F1开关.%X0 )
      P_Trig( #抽空超时沿 )
      wire#w2
      I_Contact( "触摸屏".设备配置.%X7 )
      wire#w3
      S_Coil( "触摸屏".运行错误报警F1.%X0 )
   END_RUNG
   RUNG wire#powerrail
      Contact( "中间变量".加湿阶段抽空超时报警 )
   END_RUNG wire#w1
   RUNG wire#powerrail
      Contact( "中间变量".脉动阶段抽空超时报警 )
   END_RUNG wire#w1
   RUNG wire#w2
      Contact( "触摸屏".设备配置.%X7 )
      { S7_Templates := "SrcType := Int" } EQ_Contact(in1 := "触摸屏".正使用泵的编号, in2 := 1)
   END_RUNG wire#w3
   RUNG wire#w2
      Contact( "触摸屏".设备配置.%X7 )
      { S7_Templates := "SrcType := Int" } EQ_Contact(in1 := "触摸屏".正使用泵的编号, in2 := 2)
      S_Coil( "触摸屏".运行错误报警F1.%X10 )
   END_RUNG
   // the same network as SCL:
   #_w1 := ("中间变量".预热阶段抽空超时报警 OR "中间变量".加湿阶段抽空超时报警 OR "中间变量".脉动阶段抽空超时报警) AND NOT "触摸屏".运行错误报警F1开关.%X0;
   #_w2 := #_w1 AND NOT #抽空超时沿;   // rising edge
   #抽空超时沿 := #_w1;
   IF #_w2 AND (NOT "触摸屏".设备配置.%X7 OR ("触摸屏".设备配置.%X7 AND ("触摸屏".正使用泵的编号 = 1))) THEN
       "触摸屏".运行错误报警F1.%X0 := TRUE;
   END_IF;
   IF #_w2 AND "触摸屏".设备配置.%X7 AND ("触摸屏".正使用泵的编号 = 2) THEN "触摸屏".运行错误报警F1.%X10 := TRUE; END_IF;
END_REGION

REGION Network 53: F002 回空超时
   RUNG wire#powerrail
      Contact( "中间变量".脉动阶段回空超时报警 )
      I_Contact( "触摸屏".运行错误报警F1开关.%X1 )
      S_Coil( "触摸屏".运行错误报警F1.%X1 )
   END_RUNG
   // the same network as SCL:
   IF "中间变量".脉动阶段回空超时报警 AND NOT "触摸屏".运行错误报警F1开关.%X1 THEN "触摸屏".运行错误报警F1.%X1 := TRUE; END_IF;
END_REGION

REGION Network 54: F003 保压失败
   RUNG wire#powerrail
      Contact( "中间变量".保压阶段保压超时报警 )
      I_Contact( "触摸屏".运行错误报警F1开关.%X2 )
      S_Coil( "触摸屏".运行错误报警F1.%X2 )
   END_RUNG
   // the same network as SCL:
   IF "中间变量".保压阶段保压超时报警 AND NOT "触摸屏".运行错误报警F1开关.%X2 THEN "触摸屏".运行错误报警F1.%X2 := TRUE; END_IF;
END_REGION

REGION Network 55: F004 加湿超时
   RUNG wire#powerrail
      Contact( "中间变量".加湿阶段加湿超时报警 )
      I_Contact( "触摸屏".运行错误报警F1开关.%X3 )
      S_Coil( "触摸屏".运行错误报警F1.%X3 )
   END_RUNG
   // the same network as SCL:
   IF "中间变量".加湿阶段加湿超时报警 AND NOT "触摸屏".运行错误报警F1开关.%X3 THEN "触摸屏".运行错误报警F1.%X3 := TRUE; END_IF;
END_REGION

REGION Network 56: F005 加药失败，药罐可能没有被刺破。
   RUNG wire#powerrail
      Contact( "中间变量".加药阶段加药失败报警 )
      I_Contact( "触摸屏".运行错误报警F1开关.%X4 )
      S_Coil( "触摸屏".运行错误报警F1.%X4 )
   END_RUNG
   // the same network as SCL:
   IF "中间变量".加药阶段加药失败报警 AND NOT "触摸屏".运行错误报警F1开关.%X4 THEN "触摸屏".运行错误报警F1.%X4 := TRUE; END_IF;
END_REGION

REGION Network 57: F006 进药压力过高，请检查设备。
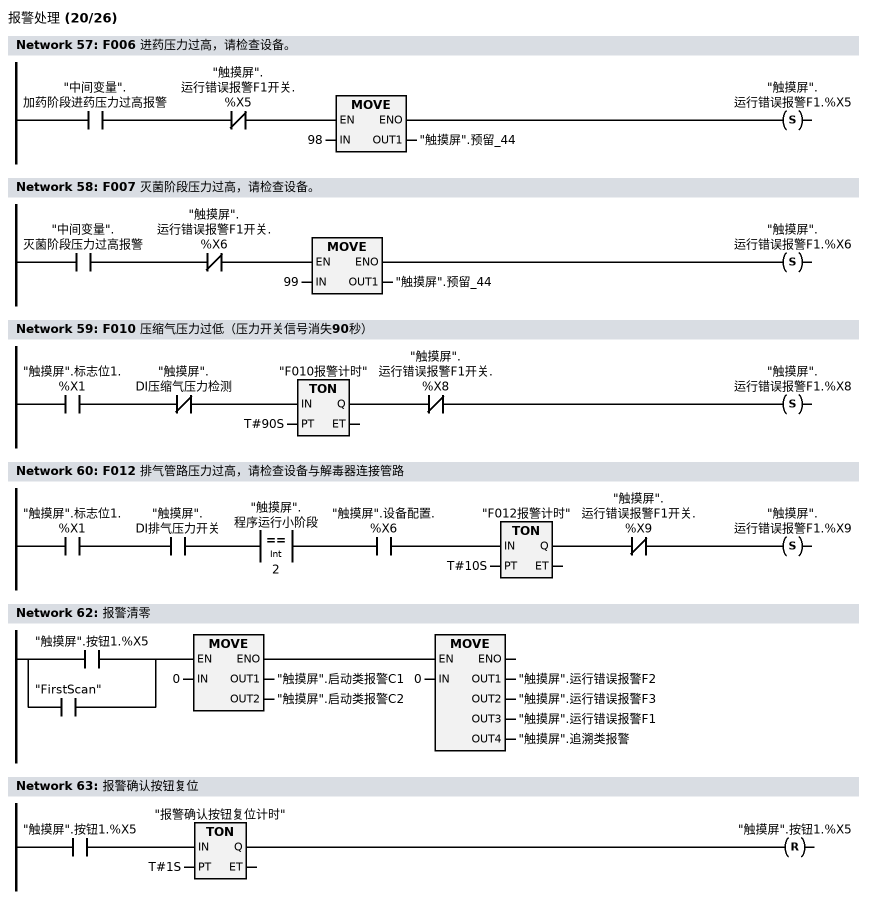
   RUNG wire#powerrail
      Contact( "中间变量".加药阶段进药压力过高报警 )
      I_Contact( "触摸屏".运行错误报警F1开关.%X5 )
      Move(in := 98, out1 => "触摸屏".预留_44)
      S_Coil( "触摸屏".运行错误报警F1.%X5 )
   END_RUNG
   // the same network as SCL:
   IF "中间变量".加药阶段进药压力过高报警 AND NOT "触摸屏".运行错误报警F1开关.%X5 THEN
       "触摸屏".预留_44 := 98;
       "触摸屏".运行错误报警F1.%X5 := TRUE;
   END_IF;
END_REGION

REGION Network 58: F007 灭菌阶段压力过高，请检查设备。
   RUNG wire#powerrail
      Contact( "中间变量".灭菌阶段压力过高报警 )
      I_Contact( "触摸屏".运行错误报警F1开关.%X6 )
      Move(in := 99, out1 => "触摸屏".预留_44)
      S_Coil( "触摸屏".运行错误报警F1.%X6 )
   END_RUNG
   // the same network as SCL:
   IF "中间变量".灭菌阶段压力过高报警 AND NOT "触摸屏".运行错误报警F1开关.%X6 THEN
       "触摸屏".预留_44 := 99;
       "触摸屏".运行错误报警F1.%X6 := TRUE;
   END_IF;
END_REGION

REGION Network 59: F010 压缩气压力过低（压力开关信号消失90秒）
   "F010报警计时".TON(IN := "触摸屏".标志位1.%X1 AND NOT "触摸屏".DI压缩气压力检测, PT := T#90S);
   IF "F010报警计时".Q AND NOT "触摸屏".运行错误报警F1开关.%X8 THEN "触摸屏".运行错误报警F1.%X8 := TRUE; END_IF;
END_REGION

REGION Network 60: F012 排气管路压力过高，请检查设备与解毒器连接管路
   "F012报警计时".TON(IN := "触摸屏".标志位1.%X1 AND "触摸屏".DI排气压力开关 AND ("触摸屏".程序运行小阶段 = 2) AND "触摸屏".设备配置.%X6,
                  PT := T#10S);
   IF "F012报警计时".Q AND NOT "触摸屏".运行错误报警F1开关.%X9 THEN "触摸屏".运行错误报警F1.%X9 := TRUE; END_IF;
END_REGION

REGION Network 61: 追溯类报警 DB48.DBW40
   // DB48.DBX40.0 W001非法条码！
   //  DB48.DBX40.1 W002请使用前门扫描枪！
   //  DB48.DBX40.2 W003请使用后门扫描枪！
   //  DB48.DBX40.3 W004重复扫描！
   //  DB48.DBX40.4 W005设备正在运行，扫描条码无效！
   //  DB48.DBX40.5 W006无此条码相关信息！
   //  DB48.DBX40.6 W007此包不能进高温灭菌器！
   //  DB48.DBX40.7 W008此包已登记为其他设备！
   //  DB48.DBX41.0 W009装载量超过90%！
   //  DB48.DBX41.1 W010有植入物，请进行生物测试！
   //  DB48.DBX41.2 W011有超大超重包，请运行超大超重程序！
   //  DB48.DBX41.3 W012此包不能进低温灭菌器！
END_REGION

REGION Network 62: 报警清零
   RUNG wire#powerrail
      Contact( "触摸屏".按钮1.%X5 )
      wire#w1
      Move(in := 0, out1 => "触摸屏".启动类报警C1, out2 => "触摸屏".启动类报警C2)
      Move(in := 0, out1 => "触摸屏".运行错误报警F2, out2 => "触摸屏".运行错误报警F3, out3 => "触摸屏".运行错误报警F1, out4 => "触摸屏".追溯类报警)
   END_RUNG
   RUNG wire#powerrail
      Contact( "FirstScan" )
   END_RUNG wire#w1
   // the same network as SCL:
   IF "触摸屏".按钮1.%X5 OR "FirstScan" THEN
       "触摸屏".启动类报警C1 := 0;
       "触摸屏".启动类报警C2 := 0;
       "触摸屏".运行错误报警F2 := 0;
       "触摸屏".运行错误报警F3 := 0;
       "触摸屏".运行错误报警F1 := 0;
       "触摸屏".追溯类报警 := 0;
   END_IF;
END_REGION

REGION Network 63: 报警确认按钮复位
   "报警确认按钮复位计时".TON(IN := "触摸屏".按钮1.%X5, PT := T#1S);
   IF "报警确认按钮复位计时".Q THEN "触摸屏".按钮1.%X5 := FALSE; END_IF;
END_REGION

REGION Network 64: 报警引发的程序退出
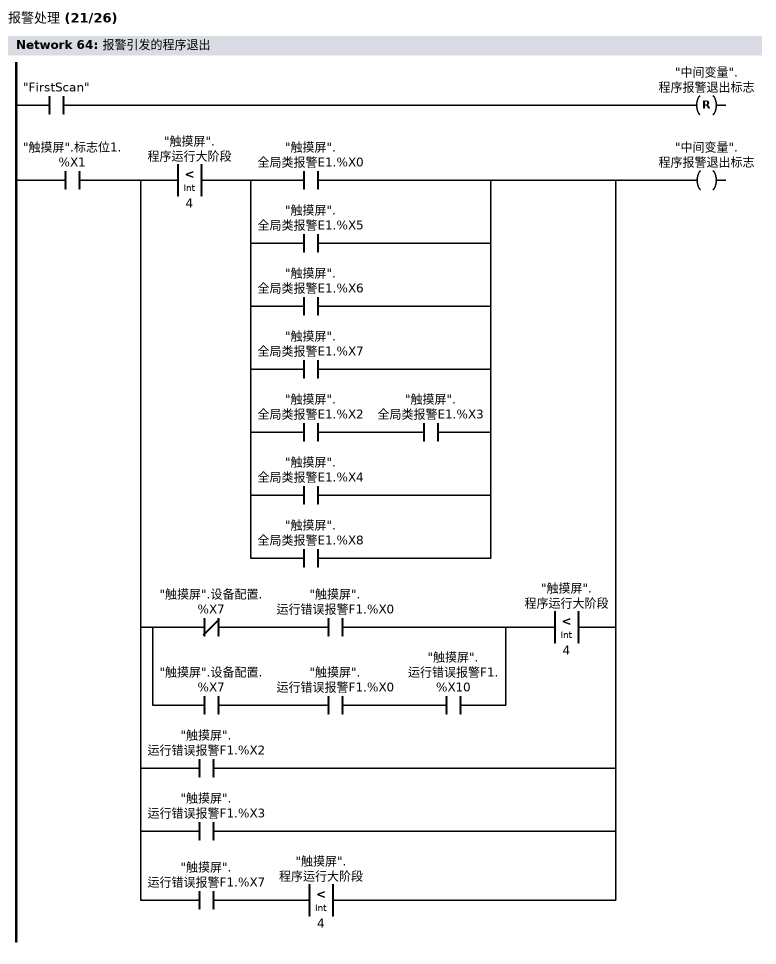
   RUNG wire#powerrail
      Contact( "FirstScan" )
      R_Coil( "中间变量".程序报警退出标志 )
   END_RUNG
   RUNG wire#powerrail
      Contact( "触摸屏".标志位1.%X1 )
      wire#w1
      { S7_Templates := "SrcType := Int" } LT_Contact(in1 := "触摸屏".程序运行大阶段, in2 := 4)
      wire#w2
      Contact( "触摸屏".全局类报警E1.%X0 )
      wire#w3
      Coil( "中间变量".程序报警退出标志 )
   END_RUNG
   RUNG wire#w2
      Contact( "触摸屏".全局类报警E1.%X5 )
   END_RUNG wire#w3
   RUNG wire#w2
      Contact( "触摸屏".全局类报警E1.%X6 )
   END_RUNG wire#w3
   RUNG wire#w2
      Contact( "触摸屏".全局类报警E1.%X7 )
   END_RUNG wire#w3
   RUNG wire#w2
      Contact( "触摸屏".全局类报警E1.%X2 )
      Contact( "触摸屏".全局类报警E1.%X3 )
   END_RUNG wire#w3
   RUNG wire#w2
      Contact( "触摸屏".全局类报警E1.%X4 )
   END_RUNG wire#w3
   RUNG wire#w2
      Contact( "触摸屏".全局类报警E1.%X8 )
   END_RUNG wire#w3
   RUNG wire#w1
      I_Contact( "触摸屏".设备配置.%X7 )
      Contact( "触摸屏".运行错误报警F1.%X0 )
      wire#w4
      { S7_Templates := "SrcType := Int" } LT_Contact(in1 := "触摸屏".程序运行大阶段, in2 := 4)
   END_RUNG wire#w3
   RUNG wire#w1
      Contact( "触摸屏".设备配置.%X7 )
      Contact( "触摸屏".运行错误报警F1.%X0 )
      Contact( "触摸屏".运行错误报警F1.%X10 )
   END_RUNG wire#w4
   RUNG wire#w1
      Contact( "触摸屏".运行错误报警F1.%X2 )
   END_RUNG wire#w3
   RUNG wire#w1
      Contact( "触摸屏".运行错误报警F1.%X3 )
   END_RUNG wire#w3
   RUNG wire#w1
      Contact( "触摸屏".运行错误报警F1.%X7 )
      { S7_Templates := "SrcType := Int" } LT_Contact(in1 := "触摸屏".程序运行大阶段, in2 := 4)
   END_RUNG wire#w3
   // the same network as SCL:
   IF "FirstScan" THEN "中间变量".程序报警退出标志 := FALSE; END_IF;
   "中间变量".程序报警退出标志 := "触摸屏".标志位1.%X1 AND ((("触摸屏".程序运行大阶段 < 4) AND ("触摸屏".全局类报警E1.%X0 OR "触摸屏".全局类报警E1.%X5 OR "触摸屏".全局类报警E1.%X6 OR "触摸屏".全局类报警E1.%X7 OR ("触摸屏".全局类报警E1.%X2 AND "触摸屏".全局类报警E1.%X3) OR "触摸屏".全局类报警E1.%X4 OR "触摸屏".全局类报警E1.%X8)) OR (((NOT "触摸屏".设备配置.%X7 AND "触摸屏".运行错误报警F1.%X0) OR ("触摸屏".设备配置.%X7 AND "触摸屏".运行错误报警F1.%X0 AND "触摸屏".运行错误报警F1.%X10)) AND ("触摸屏".程序运行大阶段 < 4)) OR "触摸屏".运行错误报警F1.%X2 OR "触摸屏".运行错误报警F1.%X3 OR ("触摸屏".运行错误报警F1.%X7 AND ("触摸屏".程序运行大阶段 < 4)));
END_REGION

REGION Network 65: 报警引发的程序暂停，可强制退出
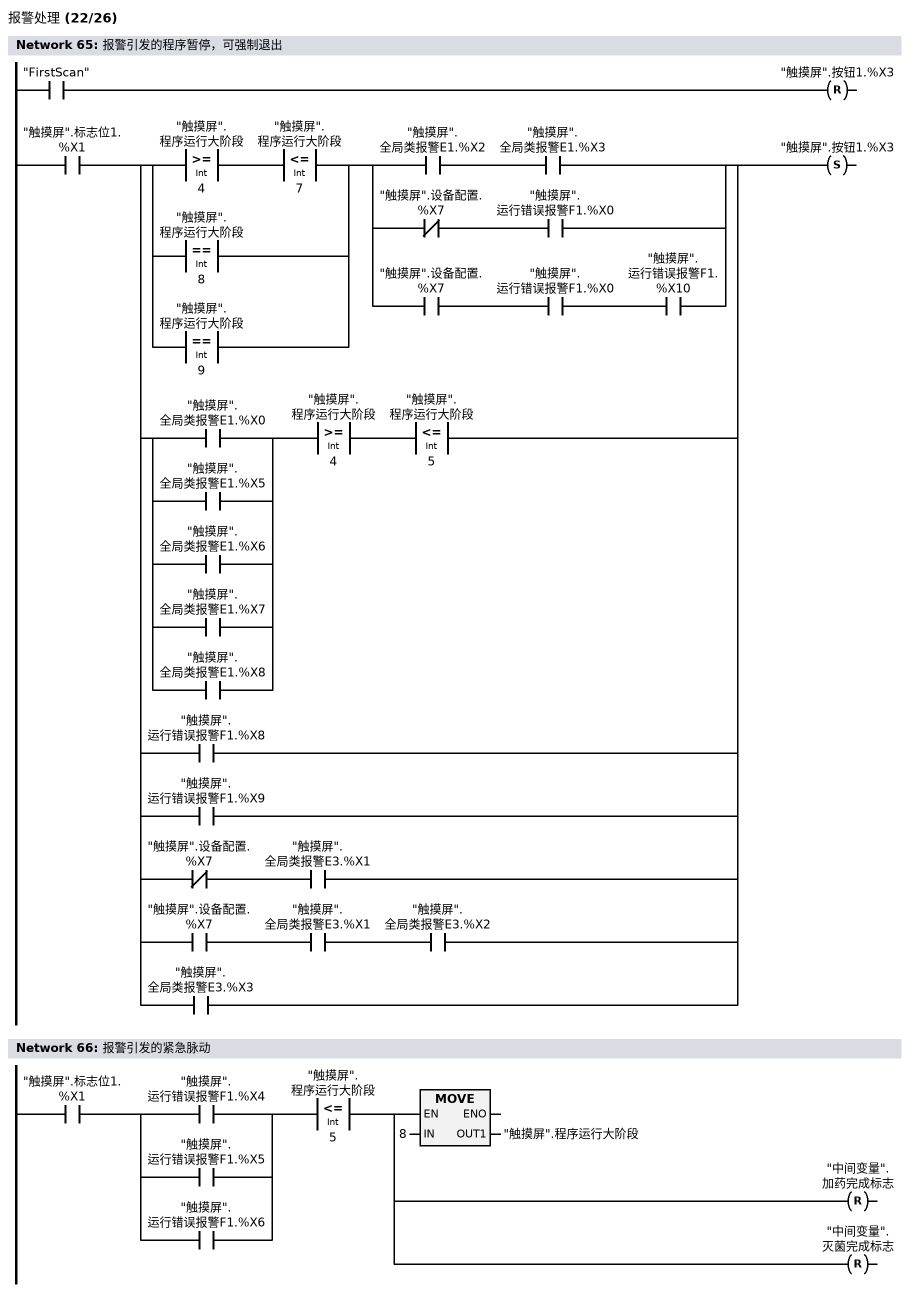
   RUNG wire#powerrail
      Contact( "FirstScan" )
      R_Coil( "触摸屏".按钮1.%X3 )
   END_RUNG
   RUNG wire#powerrail
      Contact( "触摸屏".标志位1.%X1 )
      wire#w1
      { S7_Templates := "SrcType := Int" } GE_Contact(in1 := "触摸屏".程序运行大阶段, in2 := 4)
      { S7_Templates := "SrcType := Int" } LE_Contact(in1 := "触摸屏".程序运行大阶段, in2 := 7)
      wire#w2
      Contact( "触摸屏".全局类报警E1.%X2 )
      Contact( "触摸屏".全局类报警E1.%X3 )
      wire#w3
      S_Coil( "触摸屏".按钮1.%X3 )
   END_RUNG
   RUNG wire#w1
      { S7_Templates := "SrcType := Int" } EQ_Contact(in1 := "触摸屏".程序运行大阶段, in2 := 8)
   END_RUNG wire#w2
   RUNG wire#w1
      { S7_Templates := "SrcType := Int" } EQ_Contact(in1 := "触摸屏".程序运行大阶段, in2 := 9)
   END_RUNG wire#w2
   RUNG wire#w2
      I_Contact( "触摸屏".设备配置.%X7 )
      Contact( "触摸屏".运行错误报警F1.%X0 )
   END_RUNG wire#w3
   RUNG wire#w2
      Contact( "触摸屏".设备配置.%X7 )
      Contact( "触摸屏".运行错误报警F1.%X0 )
      Contact( "触摸屏".运行错误报警F1.%X10 )
   END_RUNG wire#w3
   RUNG wire#w1
      Contact( "触摸屏".全局类报警E1.%X0 )
      wire#w4
      { S7_Templates := "SrcType := Int" } GE_Contact(in1 := "触摸屏".程序运行大阶段, in2 := 4)
      { S7_Templates := "SrcType := Int" } LE_Contact(in1 := "触摸屏".程序运行大阶段, in2 := 5)
   END_RUNG wire#w3
   RUNG wire#w1
      Contact( "触摸屏".全局类报警E1.%X5 )
   END_RUNG wire#w4
   RUNG wire#w1
      Contact( "触摸屏".全局类报警E1.%X6 )
   END_RUNG wire#w4
   RUNG wire#w1
      Contact( "触摸屏".全局类报警E1.%X7 )
   END_RUNG wire#w4
   RUNG wire#w1
      Contact( "触摸屏".全局类报警E1.%X8 )
   END_RUNG wire#w4
   RUNG wire#w1
      Contact( "触摸屏".运行错误报警F1.%X8 )
   END_RUNG wire#w3
   RUNG wire#w1
      Contact( "触摸屏".运行错误报警F1.%X9 )
   END_RUNG wire#w3
   RUNG wire#w1
      I_Contact( "触摸屏".设备配置.%X7 )
      Contact( "触摸屏".全局类报警E3.%X1 )
   END_RUNG wire#w3
   RUNG wire#w1
      Contact( "触摸屏".设备配置.%X7 )
      Contact( "触摸屏".全局类报警E3.%X1 )
      Contact( "触摸屏".全局类报警E3.%X2 )
   END_RUNG wire#w3
   RUNG wire#w1
      Contact( "触摸屏".全局类报警E3.%X3 )
   END_RUNG wire#w3
   // the same network as SCL:
   IF "FirstScan" THEN "触摸屏".按钮1.%X3 := FALSE; END_IF;
   IF "触摸屏".标志位1.%X1 AND ((((("触摸屏".程序运行大阶段 >= 4) AND ("触摸屏".程序运行大阶段 <= 7)) OR ("触摸屏".程序运行大阶段 = 8) OR ("触摸屏".程序运行大阶段 = 9)) AND (("触摸屏".全局类报警E1.%X2 AND "触摸屏".全局类报警E1.%X3) OR (NOT "触摸屏".设备配置.%X7 AND "触摸屏".运行错误报警F1.%X0) OR ("触摸屏".设备配置.%X7 AND "触摸屏".运行错误报警F1.%X0 AND "触摸屏".运行错误报警F1.%X10))) OR (("触摸屏".全局类报警E1.%X0 OR "触摸屏".全局类报警E1.%X5 OR "触摸屏".全局类报警E1.%X6 OR "触摸屏".全局类报警E1.%X7 OR "触摸屏".全局类报警E1.%X8) AND ("触摸屏".程序运行大阶段 >= 4) AND ("触摸屏".程序运行大阶段 <= 5)) OR "触摸屏".运行错误报警F1.%X8 OR "触摸屏".运行错误报警F1.%X9 OR (NOT "触摸屏".设备配置.%X7 AND "触摸屏".全局类报警E3.%X1) OR ("触摸屏".设备配置.%X7 AND "触摸屏".全局类报警E3.%X1 AND "触摸屏".全局类报警E3.%X2) OR "触摸屏".全局类报警E3.%X3) THEN
       "触摸屏".按钮1.%X3 := TRUE;
   END_IF;
END_REGION

REGION Network 66: 报警引发的紧急脉动
   RUNG wire#powerrail
      Contact( "触摸屏".标志位1.%X1 )
      wire#w1
      Contact( "触摸屏".运行错误报警F1.%X4 )
      wire#w2
      { S7_Templates := "SrcType := Int" } LE_Contact(in1 := "触摸屏".程序运行大阶段, in2 := 5)
      wire#w3
      Move(in := 8, out1 => "触摸屏".程序运行大阶段)
   END_RUNG
   RUNG wire#w1
      Contact( "触摸屏".运行错误报警F1.%X5 )
   END_RUNG wire#w2
   RUNG wire#w1
      Contact( "触摸屏".运行错误报警F1.%X6 )
   END_RUNG wire#w2
   RUNG wire#w3
      R_Coil( "中间变量".加药完成标志 )
   END_RUNG
   RUNG wire#w3
      R_Coil( "中间变量".灭菌完成标志 )
   END_RUNG
   // the same network as SCL:
   #_w1 := "触摸屏".标志位1.%X1 AND ("触摸屏".运行错误报警F1.%X4 OR "触摸屏".运行错误报警F1.%X5 OR "触摸屏".运行错误报警F1.%X6) AND ("触摸屏".程序运行大阶段 <= 5);
   IF #_w1 THEN
       "触摸屏".程序运行大阶段 := 8;
       "中间变量".加药完成标志 := FALSE;
       "中间变量".灭菌完成标志 := FALSE;
   END_IF;
END_REGION

REGION Network 67: 报警开关恢复默认
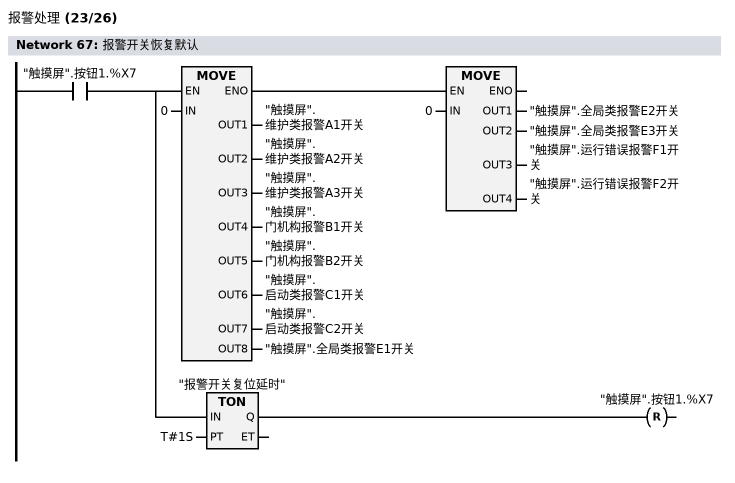
   IF "触摸屏".按钮1.%X7 THEN
       "触摸屏".维护类报警A1开关 := 0;
       "触摸屏".维护类报警A2开关 := 0;
       "触摸屏".维护类报警A3开关 := 0;
       "触摸屏".门机构报警B1开关 := 0;
       "触摸屏".门机构报警B2开关 := 0;
       "触摸屏".启动类报警C1开关 := 0;
       "触摸屏".启动类报警C2开关 := 0;
       "触摸屏".全局类报警E1开关 := 0;
       "触摸屏".全局类报警E2开关 := 0;
       "触摸屏".全局类报警E3开关 := 0;
       "触摸屏".运行错误报警F1开关 := 0;
       "触摸屏".运行错误报警F2开关 := 0;
   END_IF;
   "报警开关复位延时".TON(IN := "触摸屏".按钮1.%X7, PT := T#1S);
   IF "报警开关复位延时".Q THEN "触摸屏".按钮1.%X7 := FALSE; END_IF;
END_REGION

REGION Network 68: 设备存在报警标识
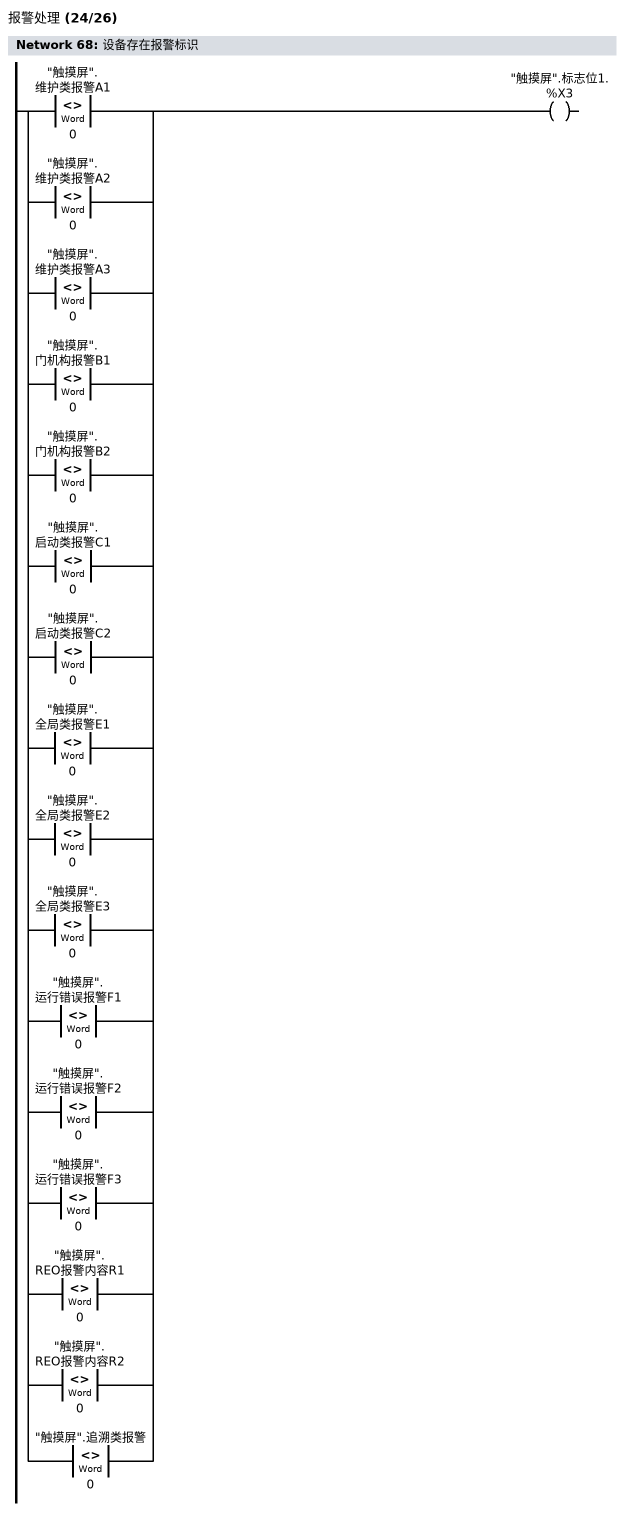
   RUNG wire#powerrail
      { S7_Templates := "SrcType := Word" } NE_Contact(in1 := "触摸屏".维护类报警A1, in2 := 0)
      wire#w1
      Coil( "触摸屏".标志位1.%X3 )
   END_RUNG
   RUNG wire#powerrail
      { S7_Templates := "SrcType := Word" } NE_Contact(in1 := "触摸屏".维护类报警A2, in2 := 0)
   END_RUNG wire#w1
   RUNG wire#powerrail
      { S7_Templates := "SrcType := Word" } NE_Contact(in1 := "触摸屏".维护类报警A3, in2 := 0)
   END_RUNG wire#w1
   RUNG wire#powerrail
      { S7_Templates := "SrcType := Word" } NE_Contact(in1 := "触摸屏".门机构报警B1, in2 := 0)
   END_RUNG wire#w1
   RUNG wire#powerrail
      { S7_Templates := "SrcType := Word" } NE_Contact(in1 := "触摸屏".门机构报警B2, in2 := 0)
   END_RUNG wire#w1
   RUNG wire#powerrail
      { S7_Templates := "SrcType := Word" } NE_Contact(in1 := "触摸屏".启动类报警C1, in2 := 0)
   END_RUNG wire#w1
   RUNG wire#powerrail
      { S7_Templates := "SrcType := Word" } NE_Contact(in1 := "触摸屏".启动类报警C2, in2 := 0)
   END_RUNG wire#w1
   RUNG wire#powerrail
      { S7_Templates := "SrcType := Word" } NE_Contact(in1 := "触摸屏".全局类报警E1, in2 := 0)
   END_RUNG wire#w1
   RUNG wire#powerrail
      { S7_Templates := "SrcType := Word" } NE_Contact(in1 := "触摸屏".全局类报警E2, in2 := 0)
   END_RUNG wire#w1
   RUNG wire#powerrail
      { S7_Templates := "SrcType := Word" } NE_Contact(in1 := "触摸屏".全局类报警E3, in2 := 0)
   END_RUNG wire#w1
   RUNG wire#powerrail
      { S7_Templates := "SrcType := Word" } NE_Contact(in1 := "触摸屏".运行错误报警F1, in2 := 0)
   END_RUNG wire#w1
   RUNG wire#powerrail
      { S7_Templates := "SrcType := Word" } NE_Contact(in1 := "触摸屏".运行错误报警F2, in2 := 0)
   END_RUNG wire#w1
   RUNG wire#powerrail
      { S7_Templates := "SrcType := Word" } NE_Contact(in1 := "触摸屏".运行错误报警F3, in2 := 0)
   END_RUNG wire#w1
   RUNG wire#powerrail
      { S7_Templates := "SrcType := Word" } NE_Contact(in1 := "触摸屏".REO报警内容R1, in2 := 0)
   END_RUNG wire#w1
   RUNG wire#powerrail
      { S7_Templates := "SrcType := Word" } NE_Contact(in1 := "触摸屏".REO报警内容R2, in2 := 0)
   END_RUNG wire#w1
   RUNG wire#powerrail
      { S7_Templates := "SrcType := Word" } NE_Contact(in1 := "触摸屏".追溯类报警, in2 := 0)
   END_RUNG wire#w1
   // the same network as SCL:
   "触摸屏".标志位1.%X3 := ("触摸屏".维护类报警A1 <> 0) OR ("触摸屏".维护类报警A2 <> 0) OR ("触摸屏".维护类报警A3 <> 0) OR ("触摸屏".门机构报警B1 <> 0) OR ("触摸屏".门机构报警B2 <> 0) OR ("触摸屏".启动类报警C1 <> 0) OR ("触摸屏".启动类报警C2 <> 0) OR ("触摸屏".全局类报警E1 <> 0) OR ("触摸屏".全局类报警E2 <> 0) OR ("触摸屏".全局类报警E3 <> 0) OR ("触摸屏".运行错误报警F1 <> 0) OR ("触摸屏".运行错误报警F2 <> 0) OR ("触摸屏".运行错误报警F3 <> 0) OR ("触摸屏".REO报警内容R1 <> 0) OR ("触摸屏".REO报警内容R2 <> 0) OR ("触摸屏".追溯类报警 <> 0);
END_REGION

REGION Network 69: 判断是否有新报警产生
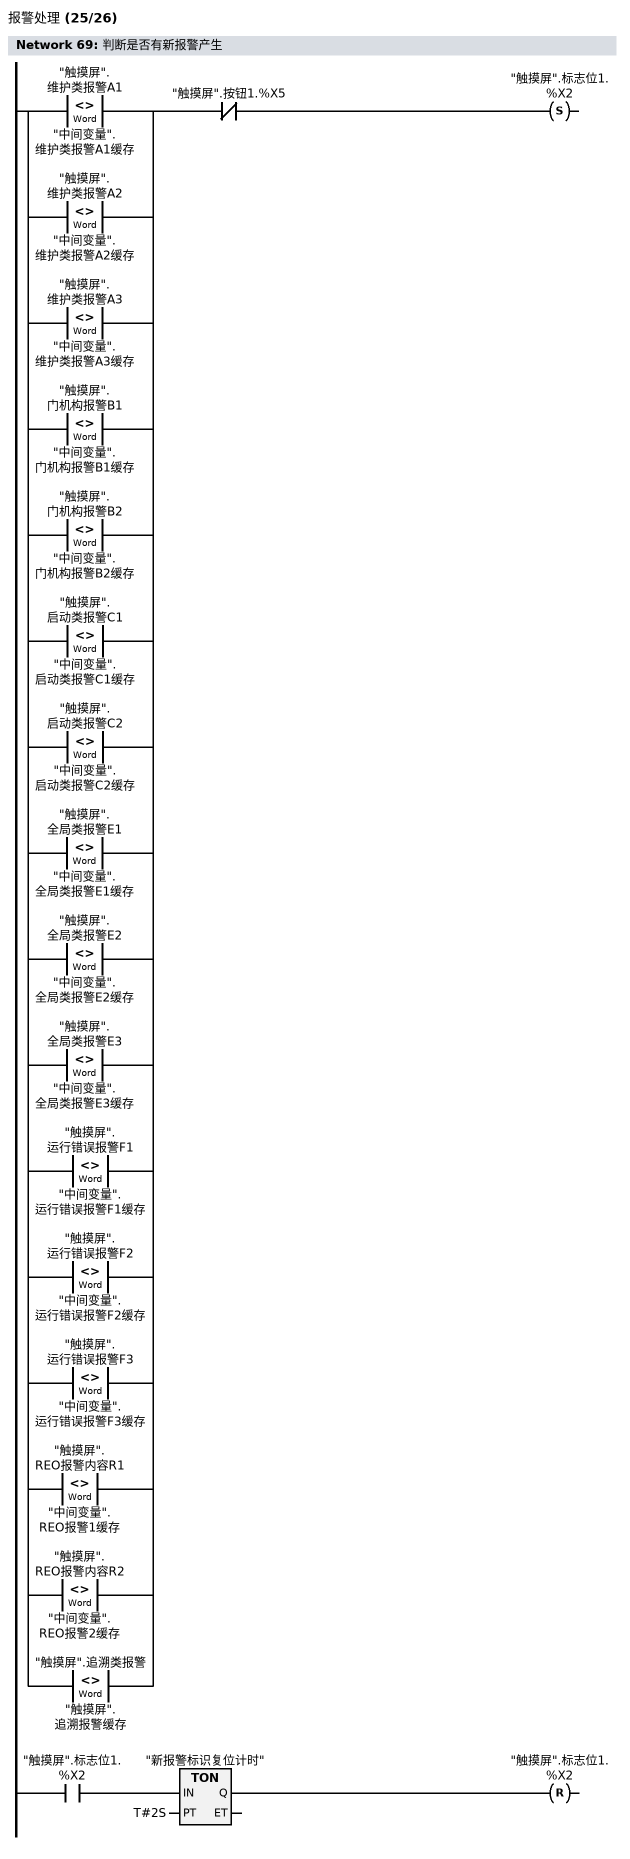
   IF (("触摸屏".维护类报警A1 <> "中间变量".维护类报警A1缓存) OR ("触摸屏".维护类报警A2 <> "中间变量".维护类报警A2缓存) OR ("触摸屏".维护类报警A3 <> "中间变量".维护类报警A3缓存) OR ("触摸屏".门机构报警B1 <> "中间变量".门机构报警B1缓存) OR ("触摸屏".门机构报警B2 <> "中间变量".门机构报警B2缓存) OR ("触摸屏".启动类报警C1 <> "中间变量".启动类报警C1缓存) OR ("触摸屏".启动类报警C2 <> "中间变量".启动类报警C2缓存) OR ("触摸屏".全局类报警E1 <> "中间变量".全局类报警E1缓存) OR ("触摸屏".全局类报警E2 <> "中间变量".全局类报警E2缓存) OR ("触摸屏".全局类报警E3 <> "中间变量".全局类报警E3缓存) OR ("触摸屏".运行错误报警F1 <> "中间变量".运行错误报警F1缓存) OR ("触摸屏".运行错误报警F2 <> "中间变量".运行错误报警F2缓存) OR ("触摸屏".运行错误报警F3 <> "中间变量".运行错误报警F3缓存) OR ("触摸屏".REO报警内容R1 <> "中间变量".REO报警1缓存) OR ("触摸屏".REO报警内容R2 <> "中间变量".REO报警2缓存) OR ("触摸屏".追溯类报警 <> "触摸屏".追溯报警缓存)) AND NOT "触摸屏".按钮1.%X5 THEN
       "触摸屏".标志位1.%X2 := TRUE;
   END_IF;
   "新报警标识复位计时".TON(IN := "触摸屏".标志位1.%X2, PT := T#2S);
   IF "新报警标识复位计时".Q THEN "触摸屏".标志位1.%X2 := FALSE; END_IF;
END_REGION

REGION Network 70: 报警信息传递给报警缓冲区
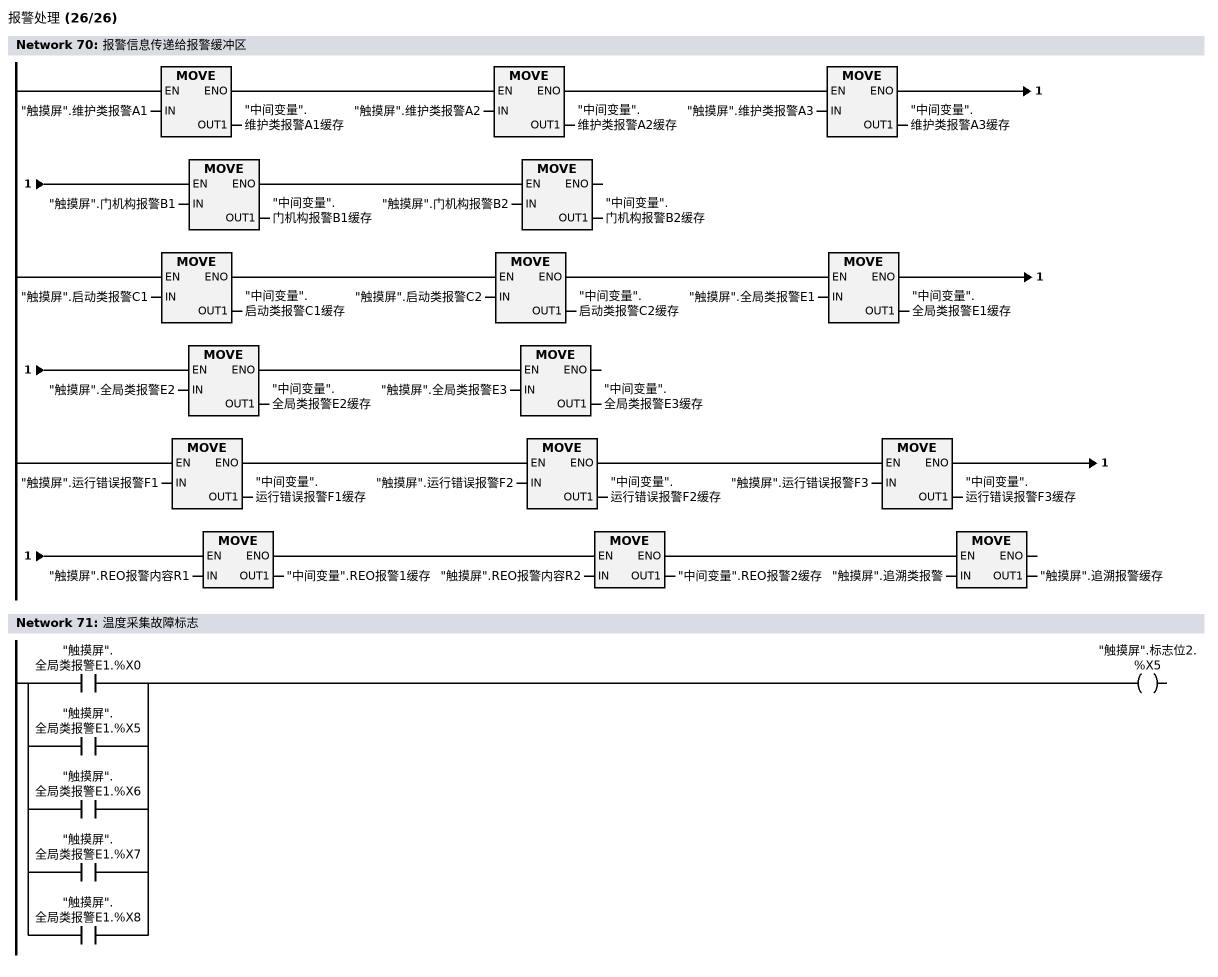
   RUNG wire#powerrail
      Move(in := "触摸屏".维护类报警A1, out1 => "中间变量".维护类报警A1缓存)
      Move(in := "触摸屏".维护类报警A2, out1 => "中间变量".维护类报警A2缓存)
      Move(in := "触摸屏".维护类报警A3, out1 => "中间变量".维护类报警A3缓存)
      Move(in := "触摸屏".门机构报警B1, out1 => "中间变量".门机构报警B1缓存)
      Move(in := "触摸屏".门机构报警B2, out1 => "中间变量".门机构报警B2缓存)
   END_RUNG
   RUNG wire#powerrail
      Move(in := "触摸屏".启动类报警C1, out1 => "中间变量".启动类报警C1缓存)
      Move(in := "触摸屏".启动类报警C2, out1 => "中间变量".启动类报警C2缓存)
      Move(in := "触摸屏".全局类报警E1, out1 => "中间变量".全局类报警E1缓存)
      Move(in := "触摸屏".全局类报警E2, out1 => "中间变量".全局类报警E2缓存)
      Move(in := "触摸屏".全局类报警E3, out1 => "中间变量".全局类报警E3缓存)
   END_RUNG
   RUNG wire#powerrail
      Move(in := "触摸屏".运行错误报警F1, out1 => "中间变量".运行错误报警F1缓存)
      Move(in := "触摸屏".运行错误报警F2, out1 => "中间变量".运行错误报警F2缓存)
      Move(in := "触摸屏".运行错误报警F3, out1 => "中间变量".运行错误报警F3缓存)
      Move(in := "触摸屏".REO报警内容R1, out1 => "中间变量".REO报警1缓存)
      Move(in := "触摸屏".REO报警内容R2, out1 => "中间变量".REO报警2缓存)
      Move(in := "触摸屏".追溯类报警, out1 => "触摸屏".追溯报警缓存)
   END_RUNG
   // the same network as SCL:
   "中间变量".维护类报警A1缓存 := "触摸屏".维护类报警A1;
   "中间变量".维护类报警A2缓存 := "触摸屏".维护类报警A2;
   "中间变量".维护类报警A3缓存 := "触摸屏".维护类报警A3;
   "中间变量".门机构报警B1缓存 := "触摸屏".门机构报警B1;
   "中间变量".门机构报警B2缓存 := "触摸屏".门机构报警B2;
   "中间变量".启动类报警C1缓存 := "触摸屏".启动类报警C1;
   "中间变量".启动类报警C2缓存 := "触摸屏".启动类报警C2;
   "中间变量".全局类报警E1缓存 := "触摸屏".全局类报警E1;
   "中间变量".全局类报警E2缓存 := "触摸屏".全局类报警E2;
   "中间变量".全局类报警E3缓存 := "触摸屏".全局类报警E3;
   "中间变量".运行错误报警F1缓存 := "触摸屏".运行错误报警F1;
   "中间变量".运行错误报警F2缓存 := "触摸屏".运行错误报警F2;
   "中间变量".运行错误报警F3缓存 := "触摸屏".运行错误报警F3;
   "中间变量".REO报警1缓存 := "触摸屏".REO报警内容R1;
   "中间变量".REO报警2缓存 := "触摸屏".REO报警内容R2;
   "触摸屏".追溯报警缓存 := "触摸屏".追溯类报警;
END_REGION

REGION Network 71: 温度采集故障标志
   RUNG wire#powerrail
      Contact( "触摸屏".全局类报警E1.%X0 )
      wire#w1
      Coil( "触摸屏".标志位2.%X5 )
   END_RUNG
   RUNG wire#powerrail
      Contact( "触摸屏".全局类报警E1.%X5 )
   END_RUNG wire#w1
   RUNG wire#powerrail
      Contact( "触摸屏".全局类报警E1.%X6 )
   END_RUNG wire#w1
   RUNG wire#powerrail
      Contact( "触摸屏".全局类报警E1.%X7 )
   END_RUNG wire#w1
   RUNG wire#powerrail
      Contact( "触摸屏".全局类报警E1.%X8 )
   END_RUNG wire#w1
   // the same network as SCL:
   "触摸屏".标志位2.%X5 := "触摸屏".全局类报警E1.%X0 OR "触摸屏".全局类报警E1.%X5 OR "触摸屏".全局类报警E1.%X6 OR "触摸屏".全局类报警E1.%X7 OR "触摸屏".全局类报警E1.%X8;
END_REGION
END_FUNCTION_BLOCK

// folder: 4网络设置

FUNCTION_BLOCK "新网络设置"   // FB28, LAD
{ S7_Optimized_Access := 'TRUE' }
VERSION : 0.1
   VAR
      强制恢复默认IP标志 : Bool;
   END_VAR
BEGIN

REGION Network 1
   // 获取当前设备IP
END_REGION

REGION Network 3: 下载程序默认IP
   // 打开前门后，按下急停按钮，再同时按下前门关位 和 前门障碍开关 持续1秒 就能恢复默认IP
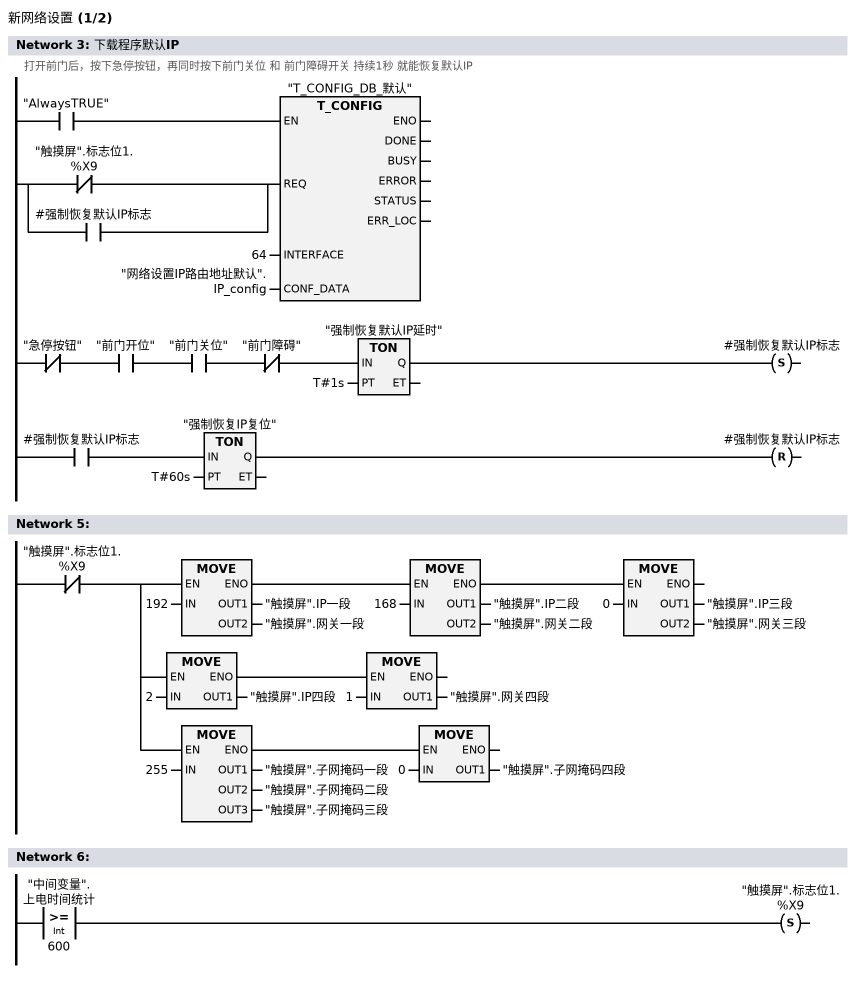
   IF "AlwaysTRUE" THEN
       "T_CONFIG_DB_默认"(Req := NOT "触摸屏".标志位1.%X9 OR #强制恢复默认IP标志,   // T_CONFIG
                        Interface := 64,
                        Conf_Data := "网络设置IP路由地址默认".IP_config);
   END_IF;
   "强制恢复默认IP延时".TON(IN := NOT "急停按钮" AND "前门开位" AND "前门关位" AND NOT "前门障碍", PT := T#1s);
   IF "强制恢复默认IP延时".Q THEN #强制恢复默认IP标志 := TRUE; END_IF;
   "强制恢复IP复位".TON(IN := #强制恢复默认IP标志, PT := T#60s);
   IF "强制恢复IP复位".Q THEN #强制恢复默认IP标志 := FALSE; END_IF;
END_REGION

REGION Network 5
   RUNG wire#powerrail
      I_Contact( "触摸屏".标志位1.%X9 )
      wire#w1
      Move(in := 192, out1 => "触摸屏".IP一段, out2 => "触摸屏".网关一段)
      Move(in := 168, out1 => "触摸屏".IP二段, out2 => "触摸屏".网关二段)
      Move(in := 0, out1 => "触摸屏".IP三段, out2 => "触摸屏".网关三段)
   END_RUNG
   RUNG wire#w1
      Move(in := 2, out1 => "触摸屏".IP四段)
      Move(in := 1, out1 => "触摸屏".网关四段)
   END_RUNG
   RUNG wire#w1
      Move(in := 255, out1 => "触摸屏".子网掩码一段, out2 => "触摸屏".子网掩码二段, out3 => "触摸屏".子网掩码三段)
      Move(in := 0, out1 => "触摸屏".子网掩码四段)
   END_RUNG
   // the same network as SCL:
   IF NOT "触摸屏".标志位1.%X9 THEN
       "触摸屏".IP一段 := 192;
       "触摸屏".网关一段 := 192;
       "触摸屏".IP二段 := 168;
       "触摸屏".网关二段 := 168;
       "触摸屏".IP三段 := 0;
       "触摸屏".网关三段 := 0;
       "触摸屏".IP四段 := 2;
       "触摸屏".网关四段 := 1;
       "触摸屏".子网掩码一段 := 255;
       "触摸屏".子网掩码二段 := 255;
       "触摸屏".子网掩码三段 := 255;
       "触摸屏".子网掩码四段 := 0;
   END_IF;
END_REGION

REGION Network 6
   RUNG wire#powerrail
      { S7_Templates := "SrcType := Int" } GE_Contact(in1 := "中间变量".上电时间统计, in2 := 600)
      S_Coil( "触摸屏".标志位1.%X9 )
   END_RUNG
   // the same network as SCL:
   IF "中间变量".上电时间统计 >= 600 THEN "触摸屏".标志位1.%X9 := TRUE; END_IF;
END_REGION

REGION Network 8: 追溯监控 IP地址与网关地址传递
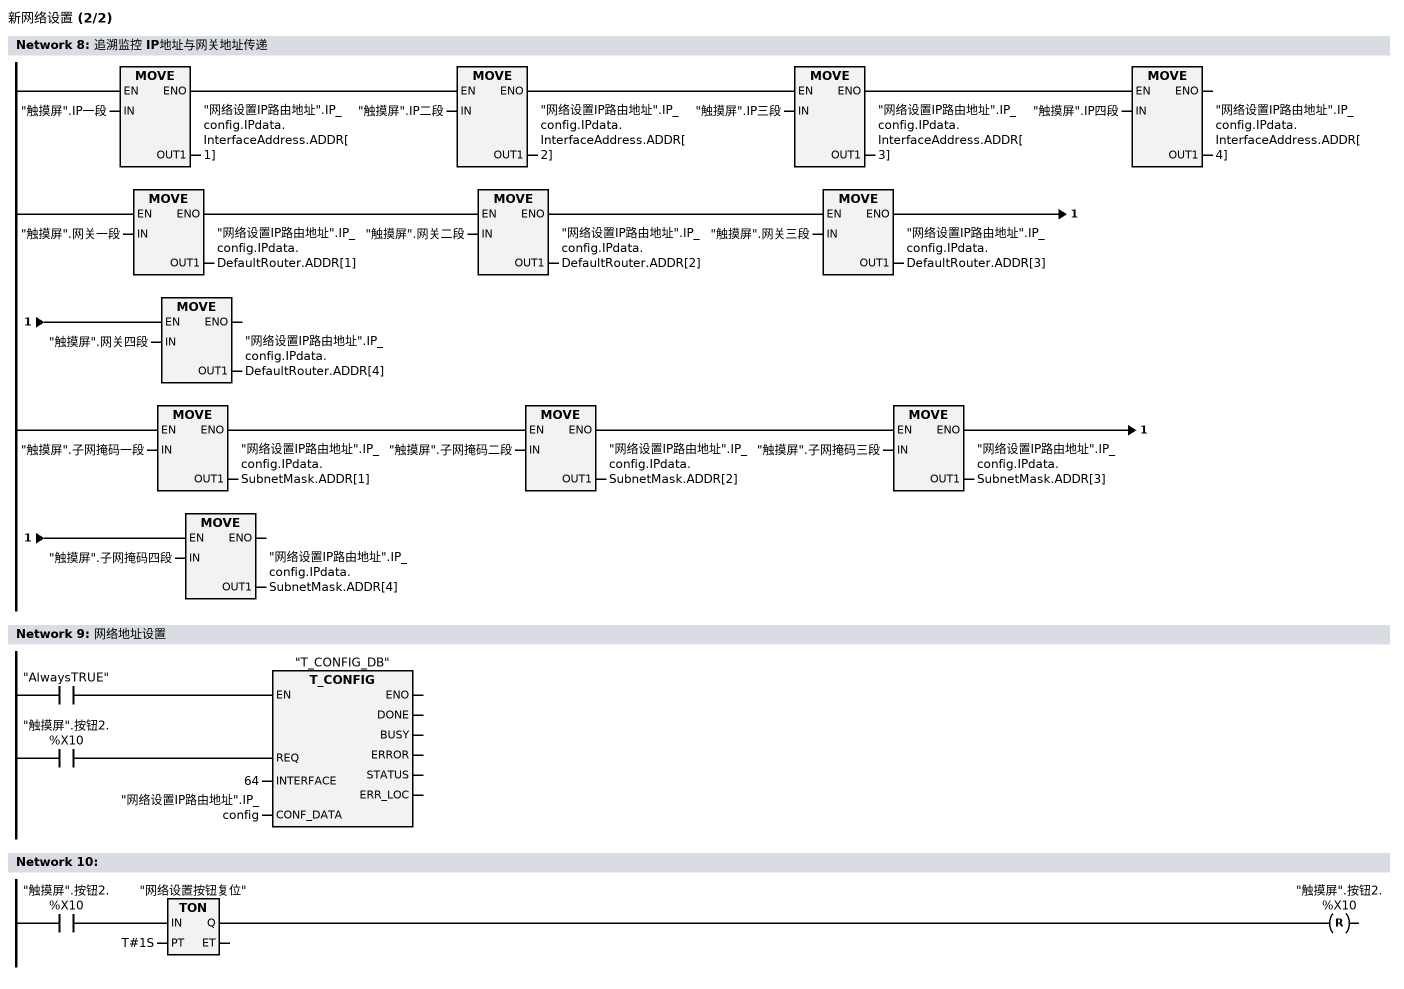
   RUNG wire#powerrail
      Move(in := "触摸屏".IP一段, out1 => "网络设置IP路由地址".IP_config.IPdata.InterfaceAddress.ADDR[1])
      Move(in := "触摸屏".IP二段, out1 => "网络设置IP路由地址".IP_config.IPdata.InterfaceAddress.ADDR[2])
      Move(in := "触摸屏".IP三段, out1 => "网络设置IP路由地址".IP_config.IPdata.InterfaceAddress.ADDR[3])
      Move(in := "触摸屏".IP四段, out1 => "网络设置IP路由地址".IP_config.IPdata.InterfaceAddress.ADDR[4])
   END_RUNG
   RUNG wire#powerrail
      Move(in := "触摸屏".网关一段, out1 => "网络设置IP路由地址".IP_config.IPdata.DefaultRouter.ADDR[1])
      Move(in := "触摸屏".网关二段, out1 => "网络设置IP路由地址".IP_config.IPdata.DefaultRouter.ADDR[2])
      Move(in := "触摸屏".网关三段, out1 => "网络设置IP路由地址".IP_config.IPdata.DefaultRouter.ADDR[3])
      Move(in := "触摸屏".网关四段, out1 => "网络设置IP路由地址".IP_config.IPdata.DefaultRouter.ADDR[4])
   END_RUNG
   RUNG wire#powerrail
      Move(in := "触摸屏".子网掩码一段, out1 => "网络设置IP路由地址".IP_config.IPdata.SubnetMask.ADDR[1])
      Move(in := "触摸屏".子网掩码二段, out1 => "网络设置IP路由地址".IP_config.IPdata.SubnetMask.ADDR[2])
      Move(in := "触摸屏".子网掩码三段, out1 => "网络设置IP路由地址".IP_config.IPdata.SubnetMask.ADDR[3])
      Move(in := "触摸屏".子网掩码四段, out1 => "网络设置IP路由地址".IP_config.IPdata.SubnetMask.ADDR[4])
   END_RUNG
   // the same network as SCL:
   "网络设置IP路由地址".IP_config.IPdata.InterfaceAddress.ADDR[1] := "触摸屏".IP一段;
   "网络设置IP路由地址".IP_config.IPdata.InterfaceAddress.ADDR[2] := "触摸屏".IP二段;
   "网络设置IP路由地址".IP_config.IPdata.InterfaceAddress.ADDR[3] := "触摸屏".IP三段;
   "网络设置IP路由地址".IP_config.IPdata.InterfaceAddress.ADDR[4] := "触摸屏".IP四段;
   "网络设置IP路由地址".IP_config.IPdata.DefaultRouter.ADDR[1] := "触摸屏".网关一段;
   "网络设置IP路由地址".IP_config.IPdata.DefaultRouter.ADDR[2] := "触摸屏".网关二段;
   "网络设置IP路由地址".IP_config.IPdata.DefaultRouter.ADDR[3] := "触摸屏".网关三段;
   "网络设置IP路由地址".IP_config.IPdata.DefaultRouter.ADDR[4] := "触摸屏".网关四段;
   "网络设置IP路由地址".IP_config.IPdata.SubnetMask.ADDR[1] := "触摸屏".子网掩码一段;
   "网络设置IP路由地址".IP_config.IPdata.SubnetMask.ADDR[2] := "触摸屏".子网掩码二段;
   "网络设置IP路由地址".IP_config.IPdata.SubnetMask.ADDR[3] := "触摸屏".子网掩码三段;
   "网络设置IP路由地址".IP_config.IPdata.SubnetMask.ADDR[4] := "触摸屏".子网掩码四段;
END_REGION

REGION Network 9: 网络地址设置
   IF "AlwaysTRUE" THEN
       "T_CONFIG_DB"(Req := "触摸屏".按钮2.%X10, Interface := 64, Conf_Data := "网络设置IP路由地址".IP_config);   // T_CONFIG
   END_IF;
END_REGION

REGION Network 10
   "网络设置按钮复位".TON(IN := "触摸屏".按钮2.%X10, PT := T#1S);
   IF "网络设置按钮复位".Q THEN "触摸屏".按钮2.%X10 := FALSE; END_IF;
END_REGION
END_FUNCTION_BLOCK

// folder: 5智慧屏功能

FUNCTION_BLOCK "智慧屏功能"   // FB23, LAD
{ S7_Optimized_Access := 'TRUE' }
VERSION : 0.1
   VAR
      沿1 : Bool;
      沿2 : Bool;
      沿3 : Bool;
      沿4 : Bool;
      冻结传递沿 : Bool;
   END_VAR
   VAR_TEMP
      各阶段打印间隔ms : DInt;
   END_VAR
   VAR_TEMP   // added for the SCL form of the ladder/FBD networks
      _w1 : Bool;
      _w2 : Bool;
      _w3 : Bool;
      _w4 : Bool;
      _w5 : Bool;
      _w6 : Bool;
      _w7 : Bool;
      _w8 : Bool;
      _w9 : Bool;
      _w10 : Bool;
      _w11 : Bool;
      _w12 : Bool;
      _w13 : Bool;
      _w14 : Bool;
      _w15 : Bool;
   END_VAR
BEGIN

REGION Network 1: 手动退出提示
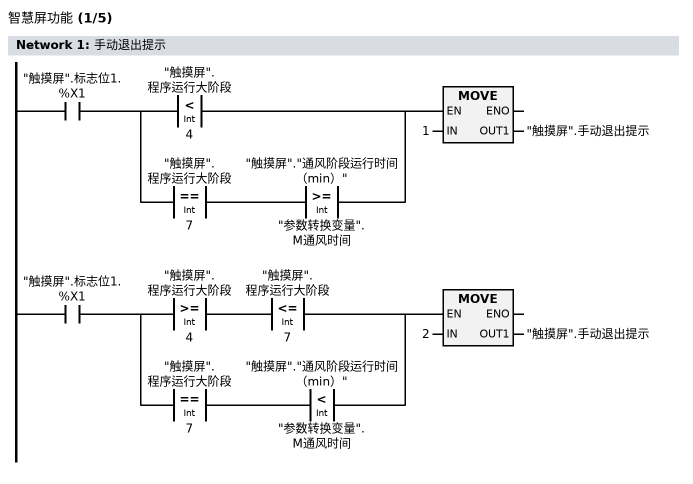
   RUNG wire#powerrail
      Contact( "触摸屏".标志位1.%X1 )
      wire#w1
      { S7_Templates := "SrcType := Int" } LT_Contact(in1 := "触摸屏".程序运行大阶段, in2 := 4)
      wire#w2
      Move(in := 1, out1 => "触摸屏".手动退出提示)
   END_RUNG
   RUNG wire#w1
      { S7_Templates := "SrcType := Int" } EQ_Contact(in1 := "触摸屏".程序运行大阶段, in2 := 7)
      { S7_Templates := "SrcType := Int" } GE_Contact(in1 := "触摸屏"."通风阶段运行时间（min）", in2 := "参数转换变量".M通风时间)
   END_RUNG wire#w2
   RUNG wire#powerrail
      Contact( "触摸屏".标志位1.%X1 )
      wire#w3
      { S7_Templates := "SrcType := Int" } GE_Contact(in1 := "触摸屏".程序运行大阶段, in2 := 4)
      { S7_Templates := "SrcType := Int" } LE_Contact(in1 := "触摸屏".程序运行大阶段, in2 := 7)
      wire#w4
      Move(in := 2, out1 => "触摸屏".手动退出提示)
   END_RUNG
   RUNG wire#w3
      { S7_Templates := "SrcType := Int" } EQ_Contact(in1 := "触摸屏".程序运行大阶段, in2 := 7)
      { S7_Templates := "SrcType := Int" } LT_Contact(in1 := "触摸屏"."通风阶段运行时间（min）", in2 := "参数转换变量".M通风时间)
   END_RUNG wire#w4
   // the same network as SCL:
   IF "触摸屏".标志位1.%X1 AND (("触摸屏".程序运行大阶段 < 4) OR (("触摸屏".程序运行大阶段 = 7) AND ("触摸屏"."通风阶段运行时间（min）" >= "参数转换变量".M通风时间))) THEN
       "触摸屏".手动退出提示 := 1;
   END_IF;
   IF "触摸屏".标志位1.%X1 AND ((("触摸屏".程序运行大阶段 >= 4) AND ("触摸屏".程序运行大阶段 <= 7)) OR (("触摸屏".程序运行大阶段 = 7) AND ("触摸屏"."通风阶段运行时间（min）" < "参数转换变量".M通风时间))) THEN
       "触摸屏".手动退出提示 := 2;
   END_IF;
END_REGION

REGION Network 2: 报表打印间隔可调
   // 20260401 韩国要求
   // "触摸屏".按钮2.%X11   打印参数默认按钮
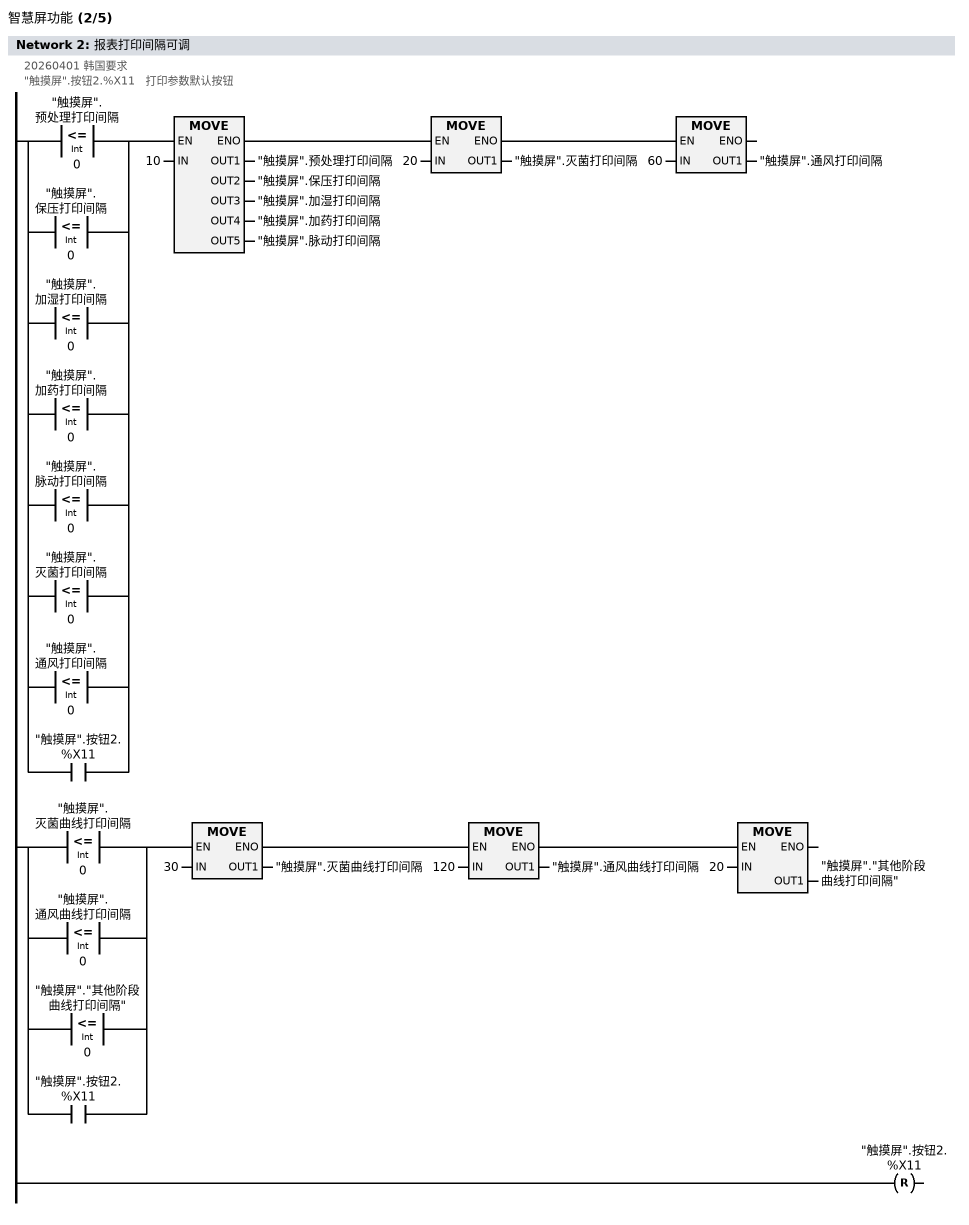
   RUNG wire#powerrail
      { S7_Templates := "SrcType := Int" } LE_Contact(in1 := "触摸屏".预处理打印间隔, in2 := 0)
      wire#w1
      Move(in := 10, out1 => "触摸屏".预处理打印间隔, out2 => "触摸屏".保压打印间隔, out3 => "触摸屏".加湿打印间隔, out4 => "触摸屏".加药打印间隔, out5 => "触摸屏".脉动打印间隔)
      Move(in := 20, out1 => "触摸屏".灭菌打印间隔)
      Move(in := 60, out1 => "触摸屏".通风打印间隔)
   END_RUNG
   RUNG wire#powerrail
      { S7_Templates := "SrcType := Int" } LE_Contact(in1 := "触摸屏".保压打印间隔, in2 := 0)
   END_RUNG wire#w1
   RUNG wire#powerrail
      { S7_Templates := "SrcType := Int" } LE_Contact(in1 := "触摸屏".加湿打印间隔, in2 := 0)
   END_RUNG wire#w1
   RUNG wire#powerrail
      { S7_Templates := "SrcType := Int" } LE_Contact(in1 := "触摸屏".加药打印间隔, in2 := 0)
   END_RUNG wire#w1
   RUNG wire#powerrail
      { S7_Templates := "SrcType := Int" } LE_Contact(in1 := "触摸屏".脉动打印间隔, in2 := 0)
   END_RUNG wire#w1
   RUNG wire#powerrail
      { S7_Templates := "SrcType := Int" } LE_Contact(in1 := "触摸屏".灭菌打印间隔, in2 := 0)
   END_RUNG wire#w1
   RUNG wire#powerrail
      { S7_Templates := "SrcType := Int" } LE_Contact(in1 := "触摸屏".通风打印间隔, in2 := 0)
   END_RUNG wire#w1
   RUNG wire#powerrail
      Contact( "触摸屏".按钮2.%X11 )
   END_RUNG wire#w1
   RUNG wire#powerrail
      { S7_Templates := "SrcType := Int" } LE_Contact(in1 := "触摸屏".灭菌曲线打印间隔, in2 := 0)
      wire#w2
      Move(in := 30, out1 => "触摸屏".灭菌曲线打印间隔)
      Move(in := 120, out1 => "触摸屏".通风曲线打印间隔)
      Move(in := 20, out1 => "触摸屏"."其他阶段 曲线打印间隔")
   END_RUNG
   RUNG wire#powerrail
      { S7_Templates := "SrcType := Int" } LE_Contact(in1 := "触摸屏".通风曲线打印间隔, in2 := 0)
   END_RUNG wire#w2
   RUNG wire#powerrail
      { S7_Templates := "SrcType := Int" } LE_Contact(in1 := "触摸屏"."其他阶段 曲线打印间隔", in2 := 0)
   END_RUNG wire#w2
   RUNG wire#powerrail
      Contact( "触摸屏".按钮2.%X11 )
   END_RUNG wire#w2
   RUNG wire#powerrail
      R_Coil( "触摸屏".按钮2.%X11 )
   END_RUNG
   // the same network as SCL:
   #_w1 := ("触摸屏".预处理打印间隔 <= 0) OR ("触摸屏".保压打印间隔 <= 0) OR ("触摸屏".加湿打印间隔 <= 0) OR ("触摸屏".加药打印间隔 <= 0) OR ("触摸屏".脉动打印间隔 <= 0) OR ("触摸屏".灭菌打印间隔 <= 0) OR ("触摸屏".通风打印间隔 <= 0) OR "触摸屏".按钮2.%X11;
   IF #_w1 THEN
       "触摸屏".预处理打印间隔 := 10;
       "触摸屏".保压打印间隔 := 10;
       "触摸屏".加湿打印间隔 := 10;
       "触摸屏".加药打印间隔 := 10;
       "触摸屏".脉动打印间隔 := 10;
       "触摸屏".灭菌打印间隔 := 20;
       "触摸屏".通风打印间隔 := 60;
   END_IF;
   #_w2 := ("触摸屏".灭菌曲线打印间隔 <= 0) OR ("触摸屏".通风曲线打印间隔 <= 0) OR ("触摸屏"."其他阶段 曲线打印间隔" <= 0) OR "触摸屏".按钮2.%X11;
   IF #_w2 THEN
       "触摸屏".灭菌曲线打印间隔 := 30;
       "触摸屏".通风曲线打印间隔 := 120;
       "触摸屏"."其他阶段 曲线打印间隔" := 20;
   END_IF;
   "触摸屏".按钮2.%X11 := FALSE;
END_REGION

REGION Network 3: 曲线打印间隔调整
